(* IEC 61131-3 sources: PLC-IsaVODE/PLC-IsaVODE/samples/plc-programs (part 5) *)

(* ---- 533-TP_1.ST ---- *)
FUNCTION UDINT_TO_TIME2:TIME

	VAR_INPUT
		IN :	UDINT;
	END_VAR

	UDINT_TO_TIME2 := DINT_TO_TIME(UDINT_TO_DINT(IN));

END_FUNCTION

FUNCTION_BLOCK T_PLC_MS_block
	VAR_OUTPUT
		T_PLC_MS :	UDINT;
	END_VAR

	VAR_EXTERNAL
		PLC_TICKS_PER_SEC :	INT;
		PLC_SYS_TICK_CNT :	DINT;
	END_VAR

	VAR
		debug :	BOOL;(*Debug-Mode ON / OFF*)
		N :	INT;(*Debug-Faktor*)
		Offset :	UDINT;(*Debug-Offset*)
		temp :	DWORD := DWORD#1;(*Debug-Offset*)
		mode :	BOOL;(*modus*)
		faktor :	UDINT;(*Systemtakt-Faktor*)
		init :	BOOL;
		v_plc_ticks_per_sec :	UDINT;
		base :	UDINT := UDINT#1000;
	END_VAR

	IF init = FALSE THEN
		v_plc_ticks_per_sec := INT_TO_UDINT(PLC_TICKS_PER_SEC);
		IF v_plc_ticks_per_sec = UDINT#1024 THEN
			faktor := UDINT#1;
			mode := FALSE;
		ELSIF v_plc_ticks_per_sec > UDINT#0 THEN
			IF v_plc_ticks_per_sec <= base THEN
				faktor := base / v_plc_ticks_per_sec;
				mode := FALSE;
			ELSE
				faktor := v_plc_ticks_per_sec / base;
				mode := TRUE;
			END_IF;
		ELSE
			faktor := UDINT#1;
		END_IF;
		init := TRUE;
	END_IF;

	IF mode THEN
		T_PLC_MS := DINT_TO_UDINT(PLC_SYS_TICK_CNT) / faktor;
	ELSE
		T_PLC_MS := DINT_TO_UDINT(PLC_SYS_TICK_CNT) * faktor;
	END_IF;

	IF debug THEN
		T_PLC_MS := (DWORD_TO_UDINT(SHL(UDINT_TO_DWORD(T_PLC_MS),N) OR SHL(temp,N)) - UDINT#1) + Offset;
	END_IF;

END_FUNCTION_BLOCK

FUNCTION_BLOCK TP_1

	VAR_INPUT
		IN :	BOOL;
		PT :	TIME;
		RST :	BOOL;
	END_VAR

	VAR_OUTPUT
		Q :	BOOL;
	END_VAR

	VAR
		tx :	TIME;
		start :	TIME;
		ix :	BOOL;
		T_PLC_MS :	T_PLC_MS_block;
	END_VAR

	T_PLC_MS();
	tx := UDINT_TO_TIME(T_PLC_MS.T_PLC_MS);

	IF RST THEN
		Q := FALSE;
	ELSIF IN AND NOT ix THEN
		Q := TRUE;
		start := tx;
	ELSIF tx - start >= PT THEN
		Q := FALSE;
	END_IF;

	ix:= IN;

END_FUNCTION_BLOCK

PROGRAM program0
  VAR
	IN :	BOOL;
	PT :	TIME;
	RST :	BOOL;
	Q :	BOOL;
	func_block : TP_1;
  END_VAR
	func_block.IN  :=IN;
	func_block.PT  :=PT;
	func_block.RST  :=RST;
	func_block();
	Q := func_block.Q;
END_PROGRAM

CONFIGURATION Config0
	VAR_GLOBAL
		PLC_TICKS_PER_SEC :	INT;
		PLC_SYS_TICK_CNT :	DINT;
	END_VAR
	RESOURCE Res0 ON PLC
		TASK task0(INTERVAL := T#20ms,PRIORITY := 0);
		PROGRAM instance0 WITH task0 : program0;
	END_RESOURCE
END_CONFIGURATION

(* ---- 534-IRTRANS_RCV_8.ST ---- *)
FUNCTION_BLOCK IRTRANS_RCV_8_Block

	VAR_INPUT
		CMD :	BOOL;
	END_VAR

	VAR_IN_OUT
		DEV :	STRING;
		KEY :	STRING;
	END_VAR

	VAR_INPUT
		DEV_CODE :	STRING;
		KEY_CODE_0 :	STRING;
		KEY_CODE_1 :	STRING;
		KEY_CODE_2 :	STRING;
		KEY_CODE_3 :	STRING;
		KEY_CODE_4 :	STRING;
		KEY_CODE_5 :	STRING;
		KEY_CODE_6 :	STRING;
		KEY_CODE_7 :	STRING;
	END_VAR

	VAR_OUTPUT
		Q0 :	BOOL;
		Q1 :	BOOL;
		Q2 :	BOOL;
		Q3 :	BOOL;
		Q4 :	BOOL;
		Q5 :	BOOL;
		Q6 :	BOOL;
		Q7 :	BOOL;
	END_VAR

	VAR
		decode :	BOOL;
	END_VAR

	decode := cmd AND EQ_STRING(dev_code,dev);

	Q0 := EQ_STRING(key,key_code_0) AND decode;
	Q1 := EQ_STRING(key,key_code_1) AND decode;
	Q2 := EQ_STRING(key,key_code_2) AND decode;
	Q3 := EQ_STRING(key,key_code_3) AND decode;
	Q4 := EQ_STRING(key,key_code_4) AND decode;
	Q5 := EQ_STRING(key,key_code_5) AND decode;
	Q6 := EQ_STRING(key,key_code_6) AND decode;
	Q7 := EQ_STRING(key,key_code_7) AND decode;

END_FUNCTION_BLOCK

PROGRAM program0
	VAR
		CMD :	BOOL;
		DEV :	STRING;
		KEY :	STRING;
		DEV_CODE :	STRING;
		KEY_CODE_0 :	STRING;
		KEY_CODE_1 :	STRING;
		KEY_CODE_2 :	STRING;
		KEY_CODE_3 :	STRING;
		KEY_CODE_4 :	STRING;
		KEY_CODE_5 :	STRING;
		KEY_CODE_6 :	STRING;
		KEY_CODE_7 :	STRING;
		Q0 :	BOOL;
		Q1 :	BOOL;
		Q2 :	BOOL;
		Q3 :	BOOL;
		Q4 :	BOOL;
		Q5 :	BOOL;
		Q6 :	BOOL;
		Q7 :	BOOL;

		func_block : IRTRANS_RCV_8_Block;
	END_VAR
	func_block.CMD := CMD;
	func_block.DEV := DEV;
	func_block.KEY := KEY;
	func_block.DEV_CODE := DEV_CODE;
	func_block.KEY_CODE_0 := KEY_CODE_0;
	func_block.KEY_CODE_1 := KEY_CODE_1;
	func_block.KEY_CODE_2 := KEY_CODE_2;
	func_block.KEY_CODE_3 := KEY_CODE_3;
	func_block.KEY_CODE_4 := KEY_CODE_4;
	func_block.KEY_CODE_5 := KEY_CODE_5;
	func_block.KEY_CODE_6 := KEY_CODE_6;
	func_block.KEY_CODE_7 := KEY_CODE_7;

	func_block();
	DEV  := func_block.DEV;
	KEY  := func_block.KEY;
	Q0  := func_block.Q0;
	Q1  := func_block.Q1;
	Q2  := func_block.Q2;
	Q3  := func_block.Q3;
	Q4  := func_block.Q4;
	Q5  := func_block.Q5;
	Q6  := func_block.Q6;
	Q7  := func_block.Q7;

END_PROGRAM

CONFIGURATION Config0

  	RESOURCE Res0 ON PLC
    	TASK task0(INTERVAL := T#20ms,PRIORITY := 0);
    	PROGRAM instance0 WITH task0 : program0;
  	END_RESOURCE

END_CONFIGURATION

(* ---- 535-TP_X.ST ---- *)
FUNCTION UDINT_TO_TIME2:TIME

	VAR_INPUT
		IN :	UDINT;
	END_VAR

	UDINT_TO_TIME2 := DINT_TO_TIME(UDINT_TO_DINT(IN));

END_FUNCTION

FUNCTION_BLOCK T_PLC_MS_block
	VAR_OUTPUT
		T_PLC_MS :	UDINT;
	END_VAR

	VAR_EXTERNAL
		PLC_TICKS_PER_SEC :	INT;
		PLC_SYS_TICK_CNT :	DINT;
	END_VAR

	VAR
		debug :	BOOL;(*Debug-Mode ON / OFF*)
		N :	INT;(*Debug-Faktor*)
		Offset :	UDINT;(*Debug-Offset*)
		temp :	DWORD := DWORD#1;(*Debug-Offset*)
		mode :	BOOL;(*modus*)
		faktor :	UDINT;(*Systemtakt-Faktor*)
		init :	BOOL;
		v_plc_ticks_per_sec :	UDINT;
		base :	UDINT := UDINT#1000;
	END_VAR

	IF init = FALSE THEN
		v_plc_ticks_per_sec := INT_TO_UDINT(PLC_TICKS_PER_SEC);
		IF v_plc_ticks_per_sec = UDINT#1024 THEN
			faktor := UDINT#1;
			mode := FALSE;
		ELSIF v_plc_ticks_per_sec > UDINT#0 THEN
			IF v_plc_ticks_per_sec <= base THEN
				faktor := base / v_plc_ticks_per_sec;
				mode := FALSE;
			ELSE
				faktor := v_plc_ticks_per_sec / base;
				mode := TRUE;
			END_IF;
		ELSE
			faktor := UDINT#1;
		END_IF;
		init := TRUE;
	END_IF;

	IF mode THEN
		T_PLC_MS := DINT_TO_UDINT(PLC_SYS_TICK_CNT) / faktor;
	ELSE
		T_PLC_MS := DINT_TO_UDINT(PLC_SYS_TICK_CNT) * faktor;
	END_IF;

	IF debug THEN
		T_PLC_MS := (DWORD_TO_UDINT(SHL(UDINT_TO_DWORD(T_PLC_MS),N) OR SHL(temp,N)) - UDINT#1) + Offset;
	END_IF;

END_FUNCTION_BLOCK

FUNCTION_BLOCK TP_X
	VAR_INPUT
		IN :	BOOL;
		PT :	TIME;
	END_VAR

	VAR_OUTPUT
		Q :	BOOL;
		ET :	TIME;
	END_VAR

	VAR
		edge :	BOOL;
		start :	TIME;
		tx :	TIME;
		T_PLC_MS :	T_PLC_MS_block;
	END_VAR

	T_PLC_MS();
	tx := UDINT_TO_TIME2(T_PLC_MS.T_PLC_MS);

	IF IN AND NOT edge THEN
		start := tx;
		Q := PT > t#0ms;
	ELSIF Q THEN
		ET := tx - start;
		IF ET >= PT THEN
			Q := FALSE;
			ET := t#0ms;
		END_IF;
	END_IF;
	edge := IN;

END_FUNCTION_BLOCK

PROGRAM program0
  VAR
	IN :	BOOL;
	PT :	TIME;
	Q :	BOOL;
	ET :	TIME;
	func_block : TP_X;
  END_VAR
	func_block.IN  :=IN;
	func_block.PT  :=PT ;
	func_block();
	Q := func_block.Q;
	ET := func_block.ET;
END_PROGRAM

CONFIGURATION Config0
	VAR_GLOBAL
		PLC_TICKS_PER_SEC :	INT;
		PLC_SYS_TICK_CNT :	DINT;
	END_VAR
	RESOURCE Res0 ON PLC
		TASK task0(INTERVAL := T#20ms,PRIORITY := 0);
		PROGRAM instance0 WITH task0 : program0;
	END_RESOURCE
END_CONFIGURATION

(* ---- 536-EXEC.ST ---- *)
FUNCTION_BLOCK EXEC_Block
	VAR_INPUT
		STR :	STRING;
	END_VAR

	VAR_OUTPUT
		EXEC :	STRING;
	END_VAR

	VAR
		pos :	INT;
		R1 :	REAL;
		R2 :	REAL;
		operator :	STRING;
		temp :	STRING;
		uppercase :	uppercase;
		trim :	trim;
		findB_num :	findB_num;
		findB_nonum :	findB_nonum;
	END_VAR

	trim(str:=str);
	temp:=trim.trim;

	uppercase(str:=temp);
	exec:=uppercase.uppercase;

	findB_nonum(str:=exec);
	pos :=findB_nonum.findB_nonum;

	IF pos > 1 THEN
	temp := LEFT(EXEC,pos-1);
	findB_num(str:=temp);
	IF findB_num.findB_num > 0 THEN
	R1 := STRING_TO_REAL(temp);
	END_IF;
	END_IF;
	temp := RIGHT(exec,LEN(exec)-pos);
	R2 := STRING_TO_REAL(temp);
	exec := LEFT(exec,pos);

	findB_num(str:=exec);
	pos :=findB_num.findB_num;
	operator := RIGHT(exec,LEN(exec) - pos);
	IF EQ_STRING(operator,'') AND LEN(str) = 0 THEN
		exec := '';
		RETURN;
	ELSIF EQ_STRING(operator,'') THEN
		exec := str;
		RETURN;
	END_IF;
	IF EQ_STRING(operator,'^') THEN
		exec := REAL_TO_STRING(EXPT(R1, R2),'%f');
	ELSIF EQ_STRING(operator,'SQRT') THEN
		exec := REAL_TO_STRING(SQRT(R2),'%f');
	ELSIF EQ_STRING(operator,'SIN') THEN
		exec := REAL_TO_STRING(SIN(r2),'%f');
	ELSIF EQ_STRING(operator,'COS') THEN
		exec := REAL_TO_STRING(COS(r2),'%f');
	ELSIF EQ_STRING(operator,'TAN') THEN
		exec := REAL_TO_STRING(TAN(R2),'%f');
	ELSIF EQ_STRING(operator,'*') THEN
		exec := REAL_TO_STRING(R1 * R2,'%f');
	ELSIF EQ_STRING(operator,'/') THEN
		IF R2 <> 0.0 THEN exec := REAL_TO_STRING(R1 / R2,'%f'); ELSE exec := 'ERROR'; END_IF;
	ELSIF EQ_STRING(operator,'+') THEN
		exec := REAL_TO_STRING(r1 + r2,'%f');
	ELSIF EQ_STRING(operator,'-') THEN
		exec := REAL_TO_STRING(r1 - r2,'%f');
	ELSE
		exec := 'ERROR';
	END_IF;
	IF EQ_STRING(EXEC,'ERROR') THEN
		RETURN;
	ELSIF FIND(EXEC,'.') = 0 THEN
		EXEC := CONCAT(EXEC, '.0');
	ELSE
	temp := RIGHT(EXEC,1);
	IF EQ_STRING(temp,'.') THEN
		EXEC := CONCAT(EXEC,'0');
	END_IF;
	END_IF;

END_FUNCTION_BLOCK

PROGRAM program0
	VAR
		STR :	STRING;

		EXEC :	STRING;

		func_block : EXEC_Block;
	END_VAR
	func_block.STR := STR;
	func_block();
	EXEC  := func_block.EXEC;
END_PROGRAM

CONFIGURATION Config0
	RESOURCE Res0 ON PLC
		TASK task0(INTERVAL := T#20ms,PRIORITY := 0);
		PROGRAM instance0 WITH task0 : program0;
	END_RESOURCE
END_CONFIGURATION

(* ---- 537-FILE_BLOCK.ST ---- *)
TYPE
  oscat_FILE_SERVER_DATA : STRUCT
	FILE_OPEN	: BOOL;
    FILENAME 	: STRING;
    MODE	 	: BYTE;
    OFFSET   	: UDINT;
    FILE_SIZE   : UDINT;
    AUTO_CLOSE	: TIME;
    ERROR	 	: BYTE;
  END_STRUCT;

  oscat_NW_BUF_LONG  : ARRAY [0..4095] OF BYTE;
  oscat_NETWORK_BUFFER :
  STRUCT
    SIZE   : UINT;
    BUFFER : oscat_NW_BUF_LONG;
  END_STRUCT;
END_TYPE

FUNCTION_BLOCK FILE_BLOCK

	VAR_IN_OUT
		MODE :	BYTE;
		FILENAME :	STRING;
		FSD :	oscat_FILE_SERVER_DATA;
		PT :	oscat_NETWORK_BUFFER;
	END_VAR

	VAR_INPUT
		POS :	UDINT;
	END_VAR

	VAR_OUTPUT
		ERROR :	BYTE;
		DATA :	BYTE;
	END_VAR

	VAR
		stepp :	INT;
		i :	INT;
		data_start :	UDINT;
		data_stop :	UDINT;
	END_VAR

	CASE stepp OF
	0:	IF MODE > BYTE#0 THEN
			ERROR := BYTE#0;
			IF FSD.FILE_OPEN AND (FSD.FILE_SIZE = UDINT#0 OR POS >= FSD.FILE_SIZE) THEN
				ERROR := BYTE#255;
				MODE := BYTE#0;
			ELSIF POS < data_start OR POS > data_stop OR NOT FSD.FILE_OPEN THEN
				FSD.FILENAME := FILENAME;
				FSD.MODE := BYTE#1;
				FSD.OFFSET := POS;
				PT.SIZE := UINT#65535;
				data_start := UDINT#0;
				data_stop := UDINT#0;
				stepp := 10;
			ELSE
				i := UDINT_TO_INT(POS - data_start);
				DATA := PT.BUFFER[i];
				MODE := BYTE#0;
			END_IF;
		END_IF;

	10:	IF FSD.MODE = BYTE#0 THEN
			IF FSD.ERROR > BYTE#0 THEN
				ERROR := FSD.ERROR;
				MODE := BYTE#0;
			ELSE
				data_start := POS;
				data_stop := POS + UINT_TO_UDINT(PT.SIZE) - UDINT#1;
			END_IF;
			stepp := 0;
		END_IF;
	END_CASE;
END_FUNCTION_BLOCK

PROGRAM program0
	VAR
		MODE :	BYTE;
		FILENAME :	STRING;
		FSD :	oscat_FILE_SERVER_DATA;
		PT :	oscat_NETWORK_BUFFER;
		POS :	UDINT;
		ERROR :	BYTE;
		DATA :	BYTE;

		func_block : FILE_BLOCK;
	END_VAR
	func_block.MODE    :=MODE    ;
	func_block.FILENAME:=FILENAME;
	func_block.FSD     :=FSD     ;
	func_block.PT      :=PT      ;
	func_block.POS     :=POS     ;
	func_block();
	MODE    := func_block.MODE    ;
	FILENAME:= func_block.FILENAME;
	FSD     := func_block.FSD     ;
	PT      := func_block.PT      ;
	ERROR   := func_block.ERROR;
	DATA    := func_block.DATA;

END_PROGRAM

CONFIGURATION Config0
  RESOURCE Res0 ON PLC
    TASK task0(INTERVAL := T#20ms,PRIORITY := 0);
    PROGRAM instance0 WITH task0 : program0;
  END_RESOURCE
END_CONFIGURATION

(* ---- 538-TMAX.ST ---- *)
FUNCTION UDINT_TO_TIME2:TIME

	VAR_INPUT
		IN :	UDINT;
	END_VAR

	UDINT_TO_TIME2 := DINT_TO_TIME(UDINT_TO_DINT(IN));

END_FUNCTION

FUNCTION_BLOCK T_PLC_MS_block
	VAR_OUTPUT
		T_PLC_MS :	UDINT;
	END_VAR

	VAR_EXTERNAL
		PLC_TICKS_PER_SEC :	INT;
		PLC_SYS_TICK_CNT :	DINT;
	END_VAR

	VAR
		debug :	BOOL;(*Debug-Mode ON / OFF*)
		N :	INT;(*Debug-Faktor*)
		Offset :	UDINT;(*Debug-Offset*)
		temp :	DWORD := DWORD#1;(*Debug-Offset*)
		mode :	BOOL;(*modus*)
		faktor :	UDINT;(*Systemtakt-Faktor*)
		init :	BOOL;
		v_plc_ticks_per_sec :	UDINT;
		base :	UDINT := UDINT#1000;
	END_VAR

	IF init = FALSE THEN
		v_plc_ticks_per_sec := INT_TO_UDINT(PLC_TICKS_PER_SEC);
		IF v_plc_ticks_per_sec = UDINT#1024 THEN
			faktor := UDINT#1;
			mode := FALSE;
		ELSIF v_plc_ticks_per_sec > UDINT#0 THEN
			IF v_plc_ticks_per_sec <= base THEN
				faktor := base / v_plc_ticks_per_sec;
				mode := FALSE;
			ELSE
				faktor := v_plc_ticks_per_sec / base;
				mode := TRUE;
			END_IF;
		ELSE
			faktor := UDINT#1;
		END_IF;
		init := TRUE;
	END_IF;

	IF mode THEN
		T_PLC_MS := DINT_TO_UDINT(PLC_SYS_TICK_CNT) / faktor;
	ELSE
		T_PLC_MS := DINT_TO_UDINT(PLC_SYS_TICK_CNT) * faktor;
	END_IF;

	IF debug THEN
		T_PLC_MS := (DWORD_TO_UDINT(SHL(UDINT_TO_DWORD(T_PLC_MS),N) OR SHL(temp,N)) - UDINT#1) + Offset;
	END_IF;

END_FUNCTION_BLOCK

FUNCTION_BLOCK TMAX

	VAR_INPUT
		IN :	BOOL;
		PT :	TIME;
	END_VAR

	VAR_OUTPUT
		Q :	BOOL;
		Z :	BOOL;
	END_VAR

	VAR
		tx :	TIME;
		start :	TIME;
		last_in :	BOOL;
		T_PLC_MS :	T_PLC_MS_block;
	END_VAR

	T_PLC_MS();
	tx:= UDINT_TO_TIME(T_PLC_MS.T_PLC_MS);

	Z := FALSE;

	IF NOT in THEN
		Q := FALSE;
	ELSIF IN AND NOT last_in THEN
		Q := TRUE;
		start := tx;
	ELSIF (tx - start >= PT) AND Q THEN
		Q := FALSE;
		Z := TRUE;
	END_IF;

	last_in := IN;

END_FUNCTION_BLOCK

PROGRAM program0
  VAR
	IN :	BOOL;
	PT :	TIME;
	Q :	BOOL;
	Z :	BOOL;
	func_block : TMAX;
  END_VAR
	func_block.IN  :=IN;
	func_block.PT  :=PT;
	func_block();
	Q := func_block.Q;
	Z := func_block.Z;

END_PROGRAM

CONFIGURATION Config0
	VAR_GLOBAL
		PLC_TICKS_PER_SEC :	INT;
		PLC_SYS_TICK_CNT :	DINT;
	END_VAR
	RESOURCE Res0 ON PLC
		TASK task0(INTERVAL := T#20ms,PRIORITY := 0);
		PROGRAM instance0 WITH task0 : program0;
	END_RESOURCE
END_CONFIGURATION

(* ---- 539-M_T.ST ---- *)
FUNCTION_BLOCK T_PLC_MS_block
	VAR_OUTPUT
		T_PLC_MS :	UDINT;
	END_VAR

	VAR_EXTERNAL
		PLC_TICKS_PER_SEC :	INT;
		PLC_SYS_TICK_CNT :	DINT;
	END_VAR

	VAR
		debug :	BOOL;(*Debug-Mode ON / OFF*)
		N :	INT;(*Debug-Faktor*)
		Offset :	UDINT;(*Debug-Offset*)
		temp :	DWORD := DWORD#1;(*Debug-Offset*)
		mode :	BOOL;(*modus*)
		faktor :	UDINT;(*Systemtakt-Faktor*)
		init :	BOOL;
		v_plc_ticks_per_sec :	UDINT;
		base :	UDINT := UDINT#1000;
	END_VAR

	IF init = FALSE THEN
		v_plc_ticks_per_sec := INT_TO_UDINT(PLC_TICKS_PER_SEC);
		IF v_plc_ticks_per_sec = UDINT#1024 THEN
			faktor := UDINT#1;
			mode := FALSE;
		ELSIF v_plc_ticks_per_sec > UDINT#0 THEN
			IF v_plc_ticks_per_sec <= base THEN
				faktor := base / v_plc_ticks_per_sec;
				mode := FALSE;
			ELSE
				faktor := v_plc_ticks_per_sec / base;
				mode := TRUE;
			END_IF;
		ELSE
			faktor := UDINT#1;
		END_IF;
		init := TRUE;
	END_IF;

	IF mode THEN
		T_PLC_MS := DINT_TO_UDINT(PLC_SYS_TICK_CNT) / faktor;
	ELSE
		T_PLC_MS := DINT_TO_UDINT(PLC_SYS_TICK_CNT) * faktor;
	END_IF;

	IF debug THEN
		T_PLC_MS := (DWORD_TO_UDINT(SHL(UDINT_TO_DWORD(T_PLC_MS),N) OR SHL(temp,N)) - UDINT#1) + Offset;
	END_IF;
END_FUNCTION_BLOCK

FUNCTION_BLOCK M_T_Block

	VAR_INPUT
		IN :	BOOL;
		TMAX :	TIME := t#10d;
		RST :	BOOL;
	END_VAR

	VAR_OUTPUT
		PT :	TIME;
		ET :	TIME;
	END_VAR

	VAR
		edge :	BOOL;
		start :	TIME;
		tx :	TIME;
		T_PLC_MS :	T_PLC_MS_Block;
	END_VAR

	(*@KEY@: WORKSHEET
	NAME: M_T
	IEC_LANGUAGE: ST
	*)
	(* read system timer *)
	T_PLC_MS();
	tx:= UDINT_TO_TIME(T_PLC_MS.T_PLC_MS);

	IF RST OR ET >= TMAX THEN
		PT := t#0s;
		ET := PT;
	ELSIF IN THEN
		IF NOT edge THEN start := tx; END_IF;
		ET := tx - start;
	ELSE
		PT := ET;
	END_IF;
	edge := IN;

END_FUNCTION_BLOCK

PROGRAM program0

	VAR
		IN :	BOOL;
		TMAX :	TIME := t#10d;
		RST :	BOOL;

		PT :	TIME;
		ET :	TIME;

		func_block : M_T_Block;
	END_VAR
	func_block.IN := IN;
	func_block.TMAX := TMAX;
	func_block.RST := RST;

	func_block();
	PT := func_block.PT;
	ET := func_block.ET;

END_PROGRAM

CONFIGURATION Config0

	VAR_GLOBAL
		PLC_TICKS_PER_SEC :	INT;
		PLC_SYS_TICK_CNT :	DINT;
	END_VAR

	RESOURCE Res0 ON PLC
		TASK task0(INTERVAL := T#20ms,PRIORITY := 0);
		PROGRAM instance0 WITH task0 : program0;
	END_RESOURCE

END_CONFIGURATION

(* ---- 540-FT_IMP.ST ---- *)
FUNCTION_BLOCK T_PLC_US_Block

	VAR_OUTPUT
		T_PLC_US :	UDINT;
	END_VAR

	VAR_EXTERNAL
		PLC_TICKS_PER_SEC :	INT;
		PLC_SYS_TICK_CNT :	DINT;
	END_VAR

	VAR
		debug :	BOOL;
		N :	INT;
		Offset :	UDINT;
		temp :	DWORD := DWORD#1;
		mode :	BOOL;
		faktor :	UDINT;
		init :	BOOL;
		v_plc_ticks_per_sec :	UDINT;
		base :	UDINT := UDINT#1000000;
	END_VAR

	IF init = FALSE THEN
		v_plc_ticks_per_sec := INT_TO_UDINT(PLC_TICKS_PER_SEC);
		IF v_plc_ticks_per_sec = UDINT#1024 THEN
			faktor := UDINT#1000;
			mode := FALSE;
		ELSIF v_plc_ticks_per_sec > UDINT#0 THEN
			IF v_plc_ticks_per_sec <= base THEN
				faktor := base / v_plc_ticks_per_sec;
				mode := FALSE;
			ELSE
				faktor := v_plc_ticks_per_sec / base;
				mode := TRUE;
			END_IF;
		ELSE
			faktor := UDINT#1;
		END_IF;
		init := TRUE;
	END_IF;

	IF mode THEN
		T_PLC_US := DINT_TO_UDINT(PLC_SYS_TICK_CNT) / faktor;
	ELSE
		T_PLC_US := DINT_TO_UDINT(PLC_SYS_TICK_CNT) * faktor;
	END_IF;

	IF debug THEN
		T_PLC_US := (DWORD_TO_UDINT(SHL(UDINT_TO_DWORD(T_PLC_US),N) OR SHL(temp,N)) - UDINT#1) + Offset;
	END_IF;

END_FUNCTION_BLOCK

FUNCTION_BLOCK FT_PT1

	VAR_INPUT
		IN :	REAL;
		T :	TIME;
		K :	REAL := 1.0;
	END_VAR

	VAR_OUTPUT
		OUT :	REAL;
	END_VAR

	VAR
		last :	UDINT;
		tx :	UDINT;
		init :	BOOL;
		T_PLC_US :	T_PLC_US_Block;
	END_VAR

	T_PLC_US();
	tx:= T_PLC_US.T_PLC_US;

	IF NOT init OR T = t#0s THEN
		init := TRUE;
		out := K * in;
	ELSE
		out := out + (in * K - out) * UDINT_TO_REAL(Tx - last) / TIME_TO_REAL(T) * 1.0E-3;
		IF ABS(out) < 1.0E-20 THEN out := 0.0; END_IF;
	END_IF;
	last := tx;

END_FUNCTION_BLOCK

FUNCTION_BLOCK FT_IMP

	VAR_INPUT
		IN :	REAL;
		T :	TIME;
		K :	REAL := 1.0;
	END_VAR

	VAR_OUTPUT
		OUT :	REAL;
	END_VAR

	VAR
		t1 :	FT_PT1;
	END_VAR

	T1(in:= in, T:=T);
	out := (in - t1.out) * K;

END_FUNCTION_BLOCK

PROGRAM program0
  VAR
	IN :	REAL;
	T :	TIME;
	K :	REAL;

	OUT :	REAL;

	func_block : FT_IMP;
  END_VAR
	func_block.IN :=IN ;
	func_block.T  :=T  ;
	func_block.K  :=K  ;
	func_block();
	OUT := func_block.OUT;
END_PROGRAM

CONFIGURATION Config0

	VAR_GLOBAL
		PLC_TICKS_PER_SEC :	INT;
		PLC_SYS_TICK_CNT :	DINT;
	END_VAR

	RESOURCE Res0 ON PLC
		TASK task0(INTERVAL := T#20ms,PRIORITY := 0);
		PROGRAM instance0 WITH task0 : program0;
	END_RESOURCE

END_CONFIGURATION

(* ---- 541-NET_VAR_BUFFER.ST ---- *)
TYPE
	oscat_aB1_64 : ARRAY[1..64] OF BYTE;
END_TYPE

TYPE

	oscat_NW_BUF_LONG  : ARRAY [0..4095] OF BYTE;

	oscat_NETWORK_BUFFER :
	STRUCT
		SIZE   : UINT;
		BUFFER : oscat_NW_BUF_LONG;
	END_STRUCT;

END_TYPE

TYPE oscat_NET_VAR_DATA :
	STRUCT
		CYCLE : UDINT;
		STATE : BYTE;
		INDEX : INT;
		ID_MAX : USINT;
		ERROR_ID : BYTE;
		BUF_SIZE : UINT;
		S_BUF : oscat_NETWORK_BUFFER;
		R_BUF : oscat_NETWORK_BUFFER;
	END_STRUCT;
END_TYPE

FUNCTION_BLOCK NET_VAR_BUFFER_Block

	VAR_OUTPUT
		ID :	BYTE;
	END_VAR

	VAR_IN_OUT
		BUF_IN :	oscat_aB1_64;
		BUF_OUT :	oscat_aB1_64;
		X :	oscat_NET_VAR_DATA;
	END_VAR

	VAR
		size :	INT;
		init :	BOOL;
		index :	INT;
		index2 :	INT;
	END_VAR

	IF NOT init THEN
		init := TRUE;
		X.ID_MAX := X.ID_MAX + USINT#1;
		ID := USINT_TO_BYTE(X.ID_MAX);
	END_IF;

	IF X.STATE > BYTE#0 AND X.ERROR_ID = BYTE#0 THEN
		index := X.index;
		IF X.STATE = BYTE#1 THEN
			size := 64;
			IF INT_TO_UINT(index + 3 + size) > X.BUF_SIZE THEN
				X.ERROR_ID := ID;
			ELSE
				X.S_BUF.BUFFER[index] := ID;
				index := index + 1;
				X.S_BUF.BUFFER[index] := BYTE#20;
				index := index + 1;
				X.S_BUF.BUFFER[index] := INT_TO_BYTE(size);
				index := index + 1;
				FOR index2 := 1 TO size DO
					X.S_BUF.BUFFER[index] := BUF_IN[index2];
					index := index + 1;
				END_FOR;
			END_IF;
		ELSIF X.STATE = BYTE#2 THEN
			index2 := index + 1;
			IF X.R_BUF.BUFFER[index] <> ID OR X.R_BUF.BUFFER[index2] <> BYTE#20 THEN
				X.ERROR_ID := ID;
			ELSE
				index := index + 2;
				size := BYTE_TO_INT(X.R_BUF.BUFFER[index]);
				index := index + 1;
				FOR index2 := 1 TO size DO
					BUF_OUT[index2] := X.R_BUF.BUFFER[index];
					index := index + 1;
				END_FOR;
			END_IF;
		END_IF;
		X.index := index;
	END_IF;

END_FUNCTION_BLOCK

PROGRAM program0
	VAR
		BUF_IN :	oscat_aB1_64;
		BUF_OUT :	oscat_aB1_64;
		X :	oscat_NET_VAR_DATA;
		ID :	BYTE;

		func_block : NET_VAR_BUFFER_Block;
	END_VAR
	func_block.BUF_IN := BUF_IN;
	func_block.BUF_OUT := BUF_OUT;
	func_block.X := X;

	func_block();
  	BUF_IN  := func_block.BUF_IN;
	BUF_OUT  := func_block.BUF_OUT;
	X  := func_block.X;
	ID  := func_block.ID;

END_PROGRAM

CONFIGURATION Config0
	RESOURCE Res0 ON PLC
		TASK task0(INTERVAL := T#20ms,PRIORITY := 0);
		PROGRAM instance0 WITH task0 : program0;
	END_RESOURCE
END_CONFIGURATION

(* ---- 542-GEN_PULSE.ST ---- *)
FUNCTION UDINT_TO_TIME2:TIME

	VAR_INPUT
		IN :	UDINT;
	END_VAR

	UDINT_TO_TIME2 := DINT_TO_TIME(UDINT_TO_DINT(IN));

END_FUNCTION

FUNCTION_BLOCK T_PLC_MS_block
	VAR_OUTPUT
		T_PLC_MS :	UDINT;
	END_VAR

	VAR_EXTERNAL
		PLC_TICKS_PER_SEC :	INT;
		PLC_SYS_TICK_CNT :	DINT;
	END_VAR

	VAR
		debug :	BOOL;(*Debug-Mode ON / OFF*)
		N :	INT;(*Debug-Faktor*)
		Offset :	UDINT;(*Debug-Offset*)
		temp :	DWORD := DWORD#1;(*Debug-Offset*)
		mode :	BOOL;(*modus*)
		faktor :	UDINT;(*Systemtakt-Faktor*)
		init :	BOOL;
		v_plc_ticks_per_sec :	UDINT;
		base :	UDINT := UDINT#1000;
	END_VAR

	IF init = FALSE THEN
		v_plc_ticks_per_sec := INT_TO_UDINT(PLC_TICKS_PER_SEC);
		IF v_plc_ticks_per_sec = UDINT#1024 THEN
			faktor := UDINT#1;
			mode := FALSE;
		ELSIF v_plc_ticks_per_sec > UDINT#0 THEN
			IF v_plc_ticks_per_sec <= base THEN
				faktor := base / v_plc_ticks_per_sec;
				mode := FALSE;
			ELSE
				faktor := v_plc_ticks_per_sec / base;
				mode := TRUE;
			END_IF;
		ELSE
			faktor := UDINT#1;
		END_IF;
		init := TRUE;
	END_IF;

	IF mode THEN
		T_PLC_MS := DINT_TO_UDINT(PLC_SYS_TICK_CNT) / faktor;
	ELSE
		T_PLC_MS := DINT_TO_UDINT(PLC_SYS_TICK_CNT) * faktor;
	END_IF;

	IF debug THEN
		T_PLC_MS := (DWORD_TO_UDINT(SHL(UDINT_TO_DWORD(T_PLC_MS),N) OR SHL(temp,N)) - UDINT#1) + Offset;
	END_IF;

END_FUNCTION_BLOCK

FUNCTION_BLOCK GEN_PULSE_Block

	VAR_INPUT
		ENQ :	BOOL := TRUE;
		PTH :	TIME;
		PTL :	TIME;
	END_VAR

	VAR_OUTPUT
		Q :	BOOL;
	END_VAR

	VAR
		T_PLC_MS :	T_PLC_MS_block;
		tx :	TIME;
		tn :	TIME;
		init :	BOOL;
	END_VAR

	IF enq THEN
		T_PLC_MS();
		tx:= UDINT_TO_TIME(T_PLC_MS.T_PLC_MS);
		IF NOT init THEN init := TRUE; tn := tx; END_IF;
		IF tx - tn >= SEL(Q, PTL, PTH) THEN
			tn := tn + SEL(Q, PTL, PTH);
			Q := NOT Q;
		END_IF;
	ELSE
		Q := FALSE;
		init := FALSE;
	END_IF;

END_FUNCTION_BLOCK

PROGRAM program0
  VAR
	ENQ :	BOOL := TRUE;
	PTH :	TIME;
	PTL :	TIME;
	Q :	BOOL;
	func_block : GEN_PULSE_Block;
  END_VAR
	func_block.ENQ  :=ENQ;
	func_block.PTH  :=PTH;
	func_block.PTL  :=PTL;
	func_block();
	Q := func_block.Q;

END_PROGRAM

CONFIGURATION Config0
	VAR_GLOBAL
		PLC_TICKS_PER_SEC :	INT;
		PLC_SYS_TICK_CNT :	DINT;
	END_VAR
	RESOURCE Res0 ON PLC
		TASK task0(INTERVAL := T#20ms,PRIORITY := 0);
		PROGRAM instance0 WITH task0 : program0;
	END_RESOURCE
END_CONFIGURATION

(* ---- 543-FT_DERIV.ST ---- *)
FUNCTION_BLOCK T_PLC_US_Block
	VAR_OUTPUT
		T_PLC_US :	UDINT;
	END_VAR

	VAR_EXTERNAL
		PLC_TICKS_PER_SEC :	INT;
		PLC_SYS_TICK_CNT :	DINT;
	END_VAR

	VAR
		debug :	BOOL;
		N :	INT;
		Offset :	UDINT;
		temp :	DWORD := DWORD#1;
		mode :	BOOL;
		faktor :	UDINT;
		init :	BOOL;
		v_plc_ticks_per_sec :	UDINT;
		base :	UDINT := UDINT#1000000;
	END_VAR

	IF init = FALSE THEN
		v_plc_ticks_per_sec := INT_TO_UDINT(PLC_TICKS_PER_SEC);
		IF v_plc_ticks_per_sec = UDINT#1024 THEN
			faktor := UDINT#1000;
			mode := FALSE;
		ELSIF v_plc_ticks_per_sec > UDINT#0 THEN
			IF v_plc_ticks_per_sec <= base THEN
				faktor := base / v_plc_ticks_per_sec;
				mode := FALSE;
			ELSE
				faktor := v_plc_ticks_per_sec / base;
				mode := TRUE;
			END_IF;
		ELSE
			faktor := UDINT#1;
		END_IF;
		init := TRUE;
	END_IF;

	IF mode THEN
		T_PLC_US := DINT_TO_UDINT(PLC_SYS_TICK_CNT) / faktor;
	ELSE
		T_PLC_US := DINT_TO_UDINT(PLC_SYS_TICK_CNT) * faktor;
	END_IF;

	IF debug THEN
		T_PLC_US := (DWORD_TO_UDINT(SHL(UDINT_TO_DWORD(T_PLC_US),N) OR SHL(temp,N)) - UDINT#1) + Offset;
	END_IF;
END_FUNCTION_BLOCK

FUNCTION_BLOCK FT_DERIV
	VAR_INPUT
		IN :	REAL;
		K :	REAL := 1.0;
		RUN :	BOOL := TRUE;
	END_VAR

	VAR_OUTPUT
		OUT :	REAL;
	END_VAR

	VAR
		old :	REAL;
		tx :	UDINT;
		last :	UDINT;
		init :	BOOL;
		tc :	REAL;
		T_PLC_US :	T_PLC_US_Block;
	END_VAR

	T_PLC_US();
	tx:= T_PLC_US.T_PLC_US;
	tc := UDINT_TO_REAL(tx - last);

	IF NOT init THEN
		init := TRUE;
		old := in;
	ELSIF run AND tc > 0.0 THEN
		out := (in - old) / tc * 1000000.0 * K;
		old := in;
	ELSE
		out := 0.0;
	END_IF;

	last := tx;

	T_PLC_US();
	tx:= T_PLC_US.T_PLC_US;

	IF NOT init THEN
		init := TRUE;
	ELSIF run AND tx - last > UDINT#0 THEN
		out := (in - old) / UDINT_TO_REAL(tx - last) * 1000000.0 * K;
	ELSE
		out := 0.0;
	END_IF;
	old := in;
	last := tx;
END_FUNCTION_BLOCK

PROGRAM program0
  VAR
	IN  :	REAL;
	K   :	REAL;
	RUN :	BOOL;

	OUT :	REAL;

	func_block : FT_DERIV;
  END_VAR
	func_block.IN :=IN ;
	func_block.K  :=K  ;
	func_block.RUN:=RUN;
	func_block();
	OUT := func_block.OUT;
END_PROGRAM

CONFIGURATION Config0
	VAR_GLOBAL
		PLC_TICKS_PER_SEC :	INT;
		PLC_SYS_TICK_CNT :	DINT;
	END_VAR

	RESOURCE Res0 ON PLC
		TASK task0(INTERVAL := T#20ms,PRIORITY := 0);
		PROGRAM instance0 WITH task0 : program0;
	END_RESOURCE
END_CONFIGURATION

(* ---- 544-REAL_TO_FRAC.ST ---- *)
TYPE oscat_FRACTION :
	STRUCT
		NUMERATOR : INT;
		DENOMINATOR : INT;
	END_STRUCT;
END_TYPE

FUNCTION_BLOCK REAL_TO_FRAC_Block

	VAR_INPUT
		X :	REAL;
		N :	INT;
	END_VAR

	VAR_OUTPUT
		REAL_TO_FRAC :	oscat_FRACTION;
	END_VAR

	VAR
		temp :	DINT;
		sign :	BOOL;
		X_gerundet :	DINT;
		X_ohne_Nachkomma :	REAL;
		Numerator :	DINT := 1;
		Denominator :	DINT := 0;
		Numerator_old :	DINT := 0;
		Denominator_old :	DINT := 1;
	END_VAR

	IF X < 0.0 THEN
		sign := TRUE;								(* Vorzeichen merken *)
		X := ABS(X);								(* Absolutwert berechnen *)
	END_IF;

	REPEAT
		X_gerundet := REAL_TO_DINT(X);

		temp := numerator * X_gerundet + numerator_old;		(* Zaehler um Vorkammawert erweitern *)
		numerator_old := numerator;							(* Zaehler der letzten Berechnung speichern *)
		numerator := temp;									(* Zaehler dieser Berechnung speichern *)

		temp := denominator * X_gerundet + denominator_old;	(* Nenner um Vorkammawert erweitern *)
		denominator_old := denominator;						(* Nenner der letzten Berechnung speichern *)
		denominator := temp;								(* Nenner dieser Berechnung speichern *)

		X_ohne_Nachkomma := DINT_TO_REAL(X_gerundet);
		IF X = X_ohne_Nachkomma THEN						(* Bruch geht ohne Rest auf *)
			IF ABS(denominator) <= INT_TO_DINT(N) THEN		(* kein Rundungsfehler *)
				numerator_old := numerator;					(* Numerator_old wird von Funktion zur�ckgegeben *)
				denominator_old := denominator;				(* Denominator_old wird von Funktion zur�ckgegeben *)
			END_IF;
			EXIT;											(* keine weitere Berechnung notwendig *)
		ELSE
			X := 1.0 / (X - X_ohne_Nachkomma);				(* Kehrwert vom Rest -> Neuer Bruch *)
		END_IF;

	UNTIL
		( ABS(Denominator) > INT_TO_DINT(N))
	END_REPEAT;

	IF sign THEN
		REAL_TO_FRAC.NUMERATOR := -1 * ABS(DINT_TO_INT(numerator_old));
	ELSE
		REAL_TO_FRAC.NUMERATOR :=  ABS(DINT_TO_INT(numerator_old));
	END_IF;

	REAL_TO_FRAC.DENOMINATOR := ABS(DINT_TO_INT(denominator_old));

END_FUNCTION_BLOCK

PROGRAM program0

	VAR
		X :	REAL;
		N :	INT;

        REAL_TO_FRAC :	oscat_FRACTION;
		func_block : REAL_TO_FRAC_Block;
	END_VAR
		func_block.X := X;
		func_block.N := N;
		func_block();
		REAL_TO_FRAC := func_block.REAL_TO_FRAC;

END_PROGRAM

CONFIGURATION Config0

	RESOURCE Res0 ON PLC
		TASK task0(INTERVAL := T#20ms,PRIORITY := 0);
		PROGRAM instance0 WITH task0 : program0;
	END_RESOURCE

END_CONFIGURATION

(* ---- 545-FT_TN8.ST ---- *)
TYPE
  	oscat_arr_0_7               : ARRAY [0..7]    OF REAL;
END_TYPE

FUNCTION_BLOCK T_PLC_MS_Block
	VAR_OUTPUT
		T_PLC_MS :	UDINT;
	END_VAR

	VAR_EXTERNAL
		PLC_TICKS_PER_SEC :	INT;
		PLC_SYS_TICK_CNT :	DINT;
	END_VAR

	VAR
		debug :	BOOL;(*Debug-Mode ON / OFF*)
		N :	INT;(*Debug-Faktor*)
		Offset :	UDINT;(*Debug-Offset*)
		temp :	DWORD := DWORD#1;(*Debug-Offset*)
		mode :	BOOL;(*modus*)
		faktor :	UDINT;(*Systemtakt-Faktor*)
		init :	BOOL;
		v_plc_ticks_per_sec :	UDINT;
		base :	UDINT := UDINT#1000;
	END_VAR

	IF init = FALSE THEN
		v_plc_ticks_per_sec := INT_TO_UDINT(PLC_TICKS_PER_SEC);
		IF v_plc_ticks_per_sec = UDINT#1024 THEN
			faktor := UDINT#1;
			mode := FALSE;
		ELSIF v_plc_ticks_per_sec > UDINT#0 THEN
			IF v_plc_ticks_per_sec <= base THEN
				faktor := base / v_plc_ticks_per_sec;
				mode := FALSE;
			ELSE
				faktor := v_plc_ticks_per_sec / base;
				mode := TRUE;
			END_IF;
		ELSE
			faktor := UDINT#1;
		END_IF;
		init := TRUE;
	END_IF;

	IF mode THEN
		T_PLC_MS := DINT_TO_UDINT(PLC_SYS_TICK_CNT) / faktor;
	ELSE
		T_PLC_MS := DINT_TO_UDINT(PLC_SYS_TICK_CNT) * faktor;
	END_IF;

	IF debug THEN
		T_PLC_MS := (DWORD_TO_UDINT(SHL(UDINT_TO_DWORD(T_PLC_MS),N) OR SHL(temp,N)) - UDINT#1) + Offset;
	END_IF;
END_FUNCTION_BLOCK

FUNCTION_BLOCK FT_TN8

	VAR_INPUT
		IN :	REAL;
		T :	TIME;
	END_VAR

	VAR_OUTPUT
		OUT :	REAL;
		TRIG :	BOOL;
	END_VAR

	VAR
		length :	INT := 8;
		X :	oscat_arr_0_7;
		cnt :	INT;
		last :	TIME;
		tx :	TIME;
		init :	BOOL;
		T_PLC_MS :	T_PLC_MS_Block;
	END_VAR

	T_PLC_MS();
	tx:= UDINT_TO_TIME(T_PLC_MS.T_PLC_MS);

	trig := FALSE;
	IF NOT init THEN
		x[cnt] := in;
		init := TRUE;
		last := tx;
	ELSIF tx - last >= (T / length) THEN
		IF cnt = length - 1 THEN cnt := 0; ELSE cnt := cnt + 1; END_IF;
		Out := X[cnt];
		x[cnt] := in;
		last := tx;
		trig := TRUE;
	END_IF;

END_FUNCTION_BLOCK

PROGRAM program0
  VAR
	IN :	REAL;
	T :	TIME;

	OUT :	REAL;
	TRIG :	BOOL;

	func_block : FT_TN8;
  END_VAR
	func_block.IN  :=IN ;
	func_block.T  :=T ;
	func_block();
	OUT := func_block.OUT;
	TRIG := func_block.TRIG;
END_PROGRAM

CONFIGURATION Config0

	VAR_GLOBAL
		PLC_TICKS_PER_SEC :	INT;
		PLC_SYS_TICK_CNT :	DINT;
	END_VAR

	RESOURCE Res0 ON PLC
		TASK task0(INTERVAL := T#20ms,PRIORITY := 0);
		PROGRAM instance0 WITH task0 : program0;
	END_RESOURCE

END_CONFIGURATION

(* ---- 546-FT_TN16.ST ---- *)
TYPE
  	oscat_arr_0_15               : ARRAY [0..15]    OF REAL;
END_TYPE

FUNCTION_BLOCK T_PLC_MS_Block
	VAR_OUTPUT
		T_PLC_MS :	UDINT;
	END_VAR

	VAR_EXTERNAL
		PLC_TICKS_PER_SEC :	INT;
		PLC_SYS_TICK_CNT :	DINT;
	END_VAR

	VAR
		debug :	BOOL;(*Debug-Mode ON / OFF*)
		N :	INT;(*Debug-Faktor*)
		Offset :	UDINT;(*Debug-Offset*)
		temp :	DWORD := DWORD#1;(*Debug-Offset*)
		mode :	BOOL;(*modus*)
		faktor :	UDINT;(*Systemtakt-Faktor*)
		init :	BOOL;
		v_plc_ticks_per_sec :	UDINT;
		base :	UDINT := UDINT#1000;
	END_VAR

	IF init = FALSE THEN
		v_plc_ticks_per_sec := INT_TO_UDINT(PLC_TICKS_PER_SEC);
		IF v_plc_ticks_per_sec = UDINT#1024 THEN
			faktor := UDINT#1;
			mode := FALSE;
		ELSIF v_plc_ticks_per_sec > UDINT#0 THEN
			IF v_plc_ticks_per_sec <= base THEN
				faktor := base / v_plc_ticks_per_sec;
				mode := FALSE;
			ELSE
				faktor := v_plc_ticks_per_sec / base;
				mode := TRUE;
			END_IF;
		ELSE
			faktor := UDINT#1;
		END_IF;
		init := TRUE;
	END_IF;

	IF mode THEN
		T_PLC_MS := DINT_TO_UDINT(PLC_SYS_TICK_CNT) / faktor;
	ELSE
		T_PLC_MS := DINT_TO_UDINT(PLC_SYS_TICK_CNT) * faktor;
	END_IF;

	IF debug THEN
		T_PLC_MS := (DWORD_TO_UDINT(SHL(UDINT_TO_DWORD(T_PLC_MS),N) OR SHL(temp,N)) - UDINT#1) + Offset;
	END_IF;
END_FUNCTION_BLOCK

FUNCTION_BLOCK FT_TN16
	VAR_INPUT
		IN :	REAL;
		T :	TIME;
	END_VAR

	VAR_OUTPUT
		OUT :	REAL;
		TRIG :	BOOL;
	END_VAR

	VAR
		length :	INT := 16;
		X :	oscat_arr_0_15;
		cnt :	INT;
		last :	TIME;
		tx :	TIME;
		init :	BOOL;
		T_PLC_MS :	T_PLC_MS_Block;
	END_VAR

	T_PLC_MS();
	tx:= UDINT_TO_TIME(T_PLC_MS.T_PLC_MS);

	trig := FALSE;
	IF NOT init THEN
		x[cnt] := in;
		init := TRUE;
		last := tx;
	ELSIF tx - last >= T / length THEN
		IF cnt = length - 1 THEN cnt := 0; ELSE cnt := cnt + 1; END_IF;
		Out := X[cnt];
		x[cnt] := in;
		last := tx;
		Trig := TRUE;
	END_IF;

END_FUNCTION_BLOCK

PROGRAM program0
  VAR
	IN :	REAL;
	T :	TIME;

	OUT :	REAL;
	TRIG :	BOOL;

	func_block : FT_TN16;
  END_VAR
	func_block.IN  :=IN ;
	func_block.T  :=T ;
	func_block();
	OUT := func_block.OUT;
	TRIG := func_block.TRIG;
END_PROGRAM

CONFIGURATION Config0

	VAR_GLOBAL
		PLC_TICKS_PER_SEC :	INT;
		PLC_SYS_TICK_CNT :	DINT;
	END_VAR

	RESOURCE Res0 ON PLC
		TASK task0(INTERVAL := T#20ms,PRIORITY := 0);
		PROGRAM instance0 WITH task0 : program0;
	END_RESOURCE

END_CONFIGURATION

(* ---- 547-FT_TN64.ST ---- *)
TYPE
	oscat_FT_TN64_array         : ARRAY [0..63]   OF REAL;
END_TYPE

FUNCTION_BLOCK T_PLC_MS_Block
	VAR_OUTPUT
		T_PLC_MS :	UDINT;
	END_VAR

	VAR_EXTERNAL
		PLC_TICKS_PER_SEC :	INT;
		PLC_SYS_TICK_CNT :	DINT;
	END_VAR

	VAR
		debug :	BOOL;(*Debug-Mode ON / OFF*)
		N :	INT;(*Debug-Faktor*)
		Offset :	UDINT;(*Debug-Offset*)
		temp :	DWORD := DWORD#1;(*Debug-Offset*)
		mode :	BOOL;(*modus*)
		faktor :	UDINT;(*Systemtakt-Faktor*)
		init :	BOOL;
		v_plc_ticks_per_sec :	UDINT;
		base :	UDINT := UDINT#1000;
	END_VAR

	IF init = FALSE THEN
		v_plc_ticks_per_sec := INT_TO_UDINT(PLC_TICKS_PER_SEC);
		IF v_plc_ticks_per_sec = UDINT#1024 THEN
			faktor := UDINT#1;
			mode := FALSE;
		ELSIF v_plc_ticks_per_sec > UDINT#0 THEN
			IF v_plc_ticks_per_sec <= base THEN
				faktor := base / v_plc_ticks_per_sec;
				mode := FALSE;
			ELSE
				faktor := v_plc_ticks_per_sec / base;
				mode := TRUE;
			END_IF;
		ELSE
			faktor := UDINT#1;
		END_IF;
		init := TRUE;
	END_IF;

	IF mode THEN
		T_PLC_MS := DINT_TO_UDINT(PLC_SYS_TICK_CNT) / faktor;
	ELSE
		T_PLC_MS := DINT_TO_UDINT(PLC_SYS_TICK_CNT) * faktor;
	END_IF;

	IF debug THEN
		T_PLC_MS := (DWORD_TO_UDINT(SHL(UDINT_TO_DWORD(T_PLC_MS),N) OR SHL(temp,N)) - UDINT#1) + Offset;
	END_IF;
END_FUNCTION_BLOCK

FUNCTION_BLOCK FT_TN64

	VAR_INPUT
		IN :	REAL;
		_T :	TIME;
	END_VAR

	VAR_OUTPUT
		OUT :	REAL;
		TRIG :	BOOL;
	END_VAR

	VAR
		length :	INT := 64;
		X :	oscat_FT_TN64_array;
		cnt :	INT;
		last :	TIME;
		tx :	TIME;
		init :	BOOL;
		T_PLC_MS :	T_PLC_MS_Block;
	END_VAR

	T_PLC_MS();
	tx:= UDINT_TO_TIME(T_PLC_MS.T_PLC_MS);

	trig := FALSE;
	IF NOT init THEN
		x[cnt] := in;
		init := TRUE;
		last := tx;
	ELSIF tx - last >= (_T / length) THEN
		IF cnt = length - 1 THEN cnt := 0; ELSE cnt := cnt + 1; END_IF;
		Out := X[cnt];
		x[cnt] := in;
		last := tx;
		trig := TRUE;
	END_IF;

END_FUNCTION_BLOCK

PROGRAM program0
  VAR
	IN :	REAL;
	_T :	TIME;

	OUT :	REAL;
	TRIG :	BOOL;

	func_block : FT_TN64;
  END_VAR
	func_block.IN  :=IN ;
	func_block._T  :=_T ;
	func_block();
	OUT := func_block.OUT;
	TRIG := func_block.TRIG;
END_PROGRAM

CONFIGURATION Config0

	VAR_GLOBAL
		PLC_TICKS_PER_SEC :	INT;
		PLC_SYS_TICK_CNT :	DINT;
	END_VAR

	RESOURCE Res0 ON PLC
		TASK task0(INTERVAL := T#20ms,PRIORITY := 0);
		PROGRAM instance0 WITH task0 : program0;
	END_RESOURCE

END_CONFIGURATION

(* ---- 548-RTC_MS.ST ---- *)
FUNCTION_BLOCK T_PLC_MS_Block
	VAR_OUTPUT
		T_PLC_MS :	UDINT;
	END_VAR

	VAR_EXTERNAL
		PLC_TICKS_PER_SEC :	INT;
		PLC_SYS_TICK_CNT :	DINT;
	END_VAR

	VAR
		debug :	BOOL;(*Debug-Mode ON / OFF*)
		N :	INT;(*Debug-Faktor*)
		Offset :	UDINT;(*Debug-Offset*)
		temp :	DWORD := DWORD#1;(*Debug-Offset*)
		mode :	BOOL;(*modus*)
		faktor :	UDINT;(*Systemtakt-Faktor*)
		init :	BOOL;
		v_plc_ticks_per_sec :	UDINT;
		base :	UDINT := UDINT#1000;
	END_VAR

	IF init = FALSE THEN
		v_plc_ticks_per_sec := INT_TO_UDINT(PLC_TICKS_PER_SEC);
		IF v_plc_ticks_per_sec = UDINT#1024 THEN
			faktor := UDINT#1;
			mode := FALSE;
		ELSIF v_plc_ticks_per_sec > UDINT#0 THEN
			IF v_plc_ticks_per_sec <= base THEN
				faktor := base / v_plc_ticks_per_sec;
				mode := FALSE;
			ELSE
				faktor := v_plc_ticks_per_sec / base;
				mode := TRUE;
			END_IF;
		ELSE
			faktor := UDINT#1;
		END_IF;
		init := TRUE;
	END_IF;

	IF mode THEN
		T_PLC_MS := DINT_TO_UDINT(PLC_SYS_TICK_CNT) / faktor;
	ELSE
		T_PLC_MS := DINT_TO_UDINT(PLC_SYS_TICK_CNT) * faktor;
	END_IF;

	IF debug THEN
		T_PLC_MS := (DWORD_TO_UDINT(SHL(UDINT_TO_DWORD(T_PLC_MS),N) OR SHL(temp,N)) - UDINT#1) + Offset;
	END_IF;
END_FUNCTION_BLOCK

FUNCTION_BLOCK RTC_MS_Block

	VAR_INPUT
		SET :	BOOL;
		SDT :	UDINT;
		SMS :	INT;
	END_VAR

	VAR_OUTPUT
		XDT :	UDINT;
		XMS :	INT;
	END_VAR

	VAR
		init :	BOOL;
		last :	UDINT;
		tx :	UDINT;
		T_PLC_MS :	T_PLC_MS_Block;
	END_VAR

	T_PLC_MS();
	tx:= T_PLC_MS.T_PLC_MS;

	IF set OR NOT init THEN
		(* clock needs to be set when set is true or after power up *)
		init := TRUE;
		xdt := SDT;
		XMS := SMS;
	ELSE
		XMS := XMS + UDINT_TO_INT(tx - last);
		(* check if one second has expired *)
		IF XMS > 999 THEN
			XDT := XDT + UDINT#1; (* add one second *)
			XMS := XMS - 1000;
		END_IF;
	END_IF;
	last := tx;

END_FUNCTION_BLOCK

PROGRAM program0

	VAR
		SET :	BOOL;
		SDT :	UDINT;
		SMS :	INT;
		XDT :	UDINT;
		XMS :	INT;
		func_block : RTC_MS_Block;
  	END_VAR
	func_block.SET  :=	SET;
	func_block.SDT  :=	SDT;
	func_block.SMS  :=	SMS;
	func_block();
	XDT := func_block.XDT;
	XMS := func_block.XMS;

END_PROGRAM

CONFIGURATION Config0

	VAR_GLOBAL
		PLC_TICKS_PER_SEC :	INT;
		PLC_SYS_TICK_CNT :	DINT;
	END_VAR

	RESOURCE Res0 ON PLC
		TASK task0(INTERVAL := T#20ms,PRIORITY := 0);
		PROGRAM instance0 WITH task0 : program0;
	END_RESOURCE

END_CONFIGURATION

(* ---- 550-CACOS.ST ---- *)
TYPE oscat_complex :
  STRUCT
	re : REAL;
	im : REAL;
  END_STRUCT;
END_TYPE

FUNCTION ATAN2:REAL
	VAR_INPUT
		X :	REAL;
		Y :	REAL;
	END_VAR

	IF X > 0.0 THEN
		ATAN2 := ATAN(Y/X);
	ELSIF X < 0.0 THEN
		IF Y >= 0.0 THEN
			ATAN2 := ATAN(Y/X) + 3.14159265358979323846264338327950288;
		ELSE
			ATAN2 := ATAN(Y/X) - 3.14159265358979323846264338327950288;
		END_IF;
	ELSIF Y > 0.0 THEN
		ATAN2 := 1.5707963267948965580;
	ELSIF Y < 0.0 THEN
		ATAN2 := -1.5707963267948965580;
	ELSE
		ATAN2 := 0.0;
	END_IF;

END_FUNCTION

FUNCTION HYPOT:REAL
	VAR_INPUT
		X :	REAL;
		Y :	REAL;
	END_VAR

	HYPOT := SQRT(x*x + y*y);
END_FUNCTION

FUNCTION_BLOCK CLOG_Block

	VAR_INPUT
		X :	oscat_complex;
	END_VAR

	VAR_OUTPUT
		CLOG :	oscat_complex;
	END_VAR

	CLOG.re := LN(HYPOT(X.re, X.im));
	CLOG.im := ATAN2(X.im, X.re);

END_FUNCTION_BLOCK

FUNCTION SGN : INT
  VAR_INPUT
    x : REAL;
  END_VAR

  IF X > 0.0 THEN
  	sgn := 1;
  ELSIF X < 0.0 THEN
  	sgn := -1;
  ELSE
  	sgn := 0;
  END_IF;
END_FUNCTION

FUNCTION_BLOCK CSQRT_Block
	VAR_INPUT
		X :	oscat_complex;
	END_VAR

	VAR_OUTPUT
		CSQRT :	oscat_complex;
	END_VAR

	VAR
		temp :	REAL;
	END_VAR

	temp := HYPOT(x.re, x.im);
	CSQRT.re :=  SQRT(0.5 * (temp + x.re));
	CSQRT.im :=  INT_TO_REAL(sgn(x.im)) * SQRT(0.5 * (temp - x.re));

END_FUNCTION_BLOCK

FUNCTION_BLOCK CACOSH_Block
	VAR_INPUT
		X :	oscat_complex;
	END_VAR

	VAR_OUTPUT
		CACOSH :	oscat_complex;
	END_VAR

	VAR
		Y :	oscat_complex;
		CLOG :	CLOG_Block;
		CSQRT :	CSQRT_Block;
	END_VAR

	y.re := (X.re - X.im)*(X.re + X.im) - 1.0;
	y.im := 2.0 * X.re * X.im;
	CSQRT(X:=y);
	y    := CSQRT.CSQRT;
	y.re := y.re + x.re;
	y.im := y.im + x.im;
	CLOG(X:=y);
	CACOSH  := CLOG.CLOG;
END_FUNCTION_BLOCK

FUNCTION_BLOCK CACOS_Block
	VAR_INPUT
		X :	oscat_complex;
	END_VAR

	VAR_OUTPUT
		CACOS :	oscat_complex;
	END_VAR

	VAR
		Y :	oscat_complex;
		CACOSH :	CACOSH_Block;
	END_VAR

	CACOSH(X:=x);
	y := CACOSH.CACOSH;
	CACOS.re := y.im;
	CACOS.im := -y.re;
END_FUNCTION_BLOCK

PROGRAM program0
  VAR
    LocalVar0 : oscat_complex;
	LocalOUT  : oscat_complex;
	func_block : CACOS_Block;
  END_VAR
	func_block.X  := LocalVar0;
	func_block();
	LocalOUT := func_block.CACOS;
END_PROGRAM

CONFIGURATION Config0
  RESOURCE Res0 ON PLC
    TASK task0(INTERVAL := T#20ms,PRIORITY := 0);
    PROGRAM instance0 WITH task0 : program0;
  END_RESOURCE
END_CONFIGURATION

(* ---- 551-NET_VAR_X8.ST ---- *)
FUNCTION_BLOCK NET_VAR_X8

	VAR_INPUT
		IN_REAL1 :	REAL;
		IN_REAL2 :	REAL;
		IN_DINT1 :	DINT;
		IN_DINT2 :	DINT;
		IN_UDINT1 :	UDINT;
		IN_UDINT2 :	UDINT;
		IN_DWORD1 :	DWORD;
		IN_DWORD2 :	DWORD;
	END_VAR

	VAR_OUTPUT
		OUT_REAL1 :	REAL;
		OUT_REAL2 :	REAL;
		OUT_DINT1 :	DINT;
		OUT_DINT2 :	DINT;
		OUT_UDINT1 :	UDINT;
		OUT_UDINT2 :	UDINT;
		OUT_DWORD1 :	DWORD;
		OUT_DWORD2 :	DWORD;
		ID :	BYTE;
	END_VAR

	VAR_IN_OUT
		X :	oscat_NET_VAR_DATA;
	END_VAR

	VAR
		init :	BOOL;
		i :	INT;
		i2 :	INT;
		index :	INT;
		index2 :	INT;
		REAL_TO_DW :	REAL_TO_DW;
		DW_TO_REAL :	DW_TO_REAL;
		ra :	oscat_nv_dw;
	END_VAR

	IF NOT init THEN
		init := TRUE;
		X.ID_MAX := X.ID_MAX + USINT#1;
		ID := USINT_TO_BYTE(X.ID_MAX);
	END_IF;

	IF X.STATE > BYTE#0 AND X.ERROR_ID = BYTE#0 THEN
		index := X.index;
		IF INT_TO_UINT(index + 34) > X.BUF_SIZE THEN
			X.ERROR_ID := ID;
		ELSE
			IF X.STATE = BYTE#1 THEN
				REAL_TO_DW(X:=IN_REAL1);
				ra[1] := REAL_TO_DW.REAL_TO_DW;
				REAL_TO_DW(X:=IN_REAL2);
				ra[2] := REAL_TO_DW.REAL_TO_DW;
				ra[3] := DINT_TO_DWORD(IN_DINT1);
				ra[4] := DINT_TO_DWORD(IN_DINT2);
				ra[5] := UDINT_TO_DWORD(IN_UDINT1);
				ra[6] := UDINT_TO_DWORD(IN_UDINT2);
				ra[7] := IN_DWORD1;
				ra[8] := IN_DWORD2;
				X.S_BUF.BUFFER[index] := ID;
				index := index + 1;
				X.S_BUF.BUFFER[index] := BYTE#21;
				index := index + 1;
				FOR i2 := 1 TO 8 DO;
					FOR i := 1 TO 4 DO;
						X.S_BUF.BUFFER[index] := DWORD_TO_BYTE(ra[i2]);
						ra[i2] := ROR(ra[i2],8);
						index := index + 1;
					END_FOR;
				END_FOR;

			ELSIF X.STATE = BYTE#2 THEN
				index2 := index + 1;
				IF X.R_BUF.BUFFER[index] <> ID OR X.R_BUF.BUFFER[index2] <> BYTE#21 THEN
					X.ERROR_ID := ID;
				ELSE
					index := index + 2;
					FOR i2 := 1 TO 8 DO;
						ra[i2] := DWORD#0;
						FOR i := 1 TO 4 DO;
							ra[i2] := ra[i2] OR BYTE_TO_DWORD(X.R_BUF.BUFFER[index]);
							ra[i2] := ROR(ra[i2],8);
							index := index + 1;
						END_FOR;
					END_FOR;
					DW_TO_REAL(X:=ra[1]);
					OUT_REAL1 := DW_TO_REAL.DW_TO_REAL;
					DW_TO_REAL(X:=ra[2]);
					OUT_REAL2 := DW_TO_REAL.DW_TO_REAL;
					OUT_DINT1 := DWORD_TO_DINT(ra[3]);
					OUT_DINT2 := DWORD_TO_DINT(ra[4]);
					OUT_UDINT1 := DWORD_TO_UDINT(ra[5]);
					OUT_UDINT2 := DWORD_TO_UDINT(ra[6]);
					OUT_DWORD1 := ra[7];
					OUT_DWORD2 := ra[8];
				END_IF;
			END_IF;
			X.index := index;
		END_IF;
	END_IF;

END_FUNCTION_BLOCK

(* ---- 552-CASIN.ST ---- *)
TYPE oscat_complex :
  STRUCT
	re : REAL;
	im : REAL;
  END_STRUCT;
END_TYPE

FUNCTION ATAN2:REAL
	VAR_INPUT
		X :	REAL;
		Y :	REAL;
	END_VAR

	IF X > 0.0 THEN
		ATAN2 := ATAN(Y/X);
	ELSIF X < 0.0 THEN
		IF Y >= 0.0 THEN
			ATAN2 := ATAN(Y/X) + 3.14159265358979323846264338327950288;
		ELSE
			ATAN2 := ATAN(Y/X) - 3.14159265358979323846264338327950288;
		END_IF;
	ELSIF Y > 0.0 THEN
		ATAN2 := 1.5707963267948965580;
	ELSIF Y < 0.0 THEN
		ATAN2 := -1.5707963267948965580;
	ELSE
		ATAN2 := 0.0;
	END_IF;

END_FUNCTION

FUNCTION HYPOT:REAL
	VAR_INPUT
		X :	REAL;
		Y :	REAL;
	END_VAR

	HYPOT := SQRT(x*x + y*y);
END_FUNCTION

FUNCTION_BLOCK CLOG_Block

	VAR_INPUT
		X :	oscat_complex;
	END_VAR

	VAR_OUTPUT
		CLOG :	oscat_complex;
	END_VAR

	CLOG.re := LN(HYPOT(X.re, X.im));
	CLOG.im := ATAN2(X.im, X.re);

END_FUNCTION_BLOCK

FUNCTION SGN : INT
  VAR_INPUT
    x : REAL;
  END_VAR

  IF X > 0.0 THEN
  	sgn := 1;
  ELSIF X < 0.0 THEN
  	sgn := -1;
  ELSE
  	sgn := 0;
  END_IF;
END_FUNCTION

FUNCTION_BLOCK CSQRT_Block
	VAR_INPUT
		X :	oscat_complex;
	END_VAR

	VAR_OUTPUT
		CSQRT :	oscat_complex;
	END_VAR

	VAR
		temp :	REAL;
	END_VAR

	temp := HYPOT(x.re, x.im);
	CSQRT.re :=  SQRT(0.5 * (temp + x.re));
	CSQRT.im :=  INT_TO_REAL(sgn(x.im)) * SQRT(0.5 * (temp - x.re));

END_FUNCTION_BLOCK

FUNCTION_BLOCK CASINH_Block
	VAR_INPUT
		X :	oscat_complex;
	END_VAR

	VAR_OUTPUT
		CASINH :	oscat_complex;
	END_VAR

	VAR
		Y :	oscat_complex;
		CLOG :	CLOG_Block;
		CSQRT :	CSQRT_Block;
	END_VAR

	y.re := (X.re - X.im)*(X.re + X.im) + 1.0;
	y.im := 2.0 * X.re * X.im;
	CSQRT(X:=y);
	y    := CSQRT.CSQRT;
	y.re := y.re + x.re;
	y.im := y.im + x.im;
	CLOG(X:=y);
	CASINH  := CLOG.CLOG;
END_FUNCTION_BLOCK

FUNCTION_BLOCK CASIN_Block
	VAR_INPUT
		X :	oscat_complex;
	END_VAR

	VAR_OUTPUT
		CASIN :	oscat_complex;
	END_VAR

	VAR
		Y :	oscat_complex;
		CASINH :	CASINH_Block;
	END_VAR

	y.re := -x.im;
	y.im := x.re;
	CASINH(X:=y);
	y := CASINH.CASINH;
	CASIN.re := y.im;
	CASIN.im := -y.re;
END_FUNCTION_BLOCK

PROGRAM program0
  VAR
    LocalVar0 : oscat_complex;
	LocalOUT  : oscat_complex;
	func_block : CASIN_Block;
  END_VAR
	func_block.X  := LocalVar0;
	func_block();
	LocalOUT := func_block.CASIN;
END_PROGRAM

CONFIGURATION Config0
  RESOURCE Res0 ON PLC
    TASK task0(INTERVAL := T#20ms,PRIORITY := 0);
    PROGRAM instance0 WITH task0 : program0;
  END_RESOURCE
END_CONFIGURATION

(* ---- 553-STRING_TO_TIME.ST ---- *)
FUNCTION_BLOCK UPPERCASE_Block

	VAR_INPUT
		STR :	STRING;
	END_VAR

	VAR_OUTPUT
		UPPERCASE :	STRING;
	END_VAR

	VAR
		char :	BYTE;
		char2 :	BYTE;
		pos :	INT;
		l :	INT;
		str_temp :	STRING;
	END_VAR

	UPPERCASE := str;
	l := LEN(str);
	FOR pos := 1 TO l DO
		char := INT_TO_BYTE(GET_CHAR(str,pos));
		char2 := TO_UPPER(char);
		IF char <> char2 THEN
			str_temp := UPPERCASE;
			UPPERCASE := REPLACE(str_temp,BYTE_TO_STRING(char2,'%c'),1,pos);
		END_IF;
	END_FOR;

END_FUNCTION_BLOCK

FUNCTION_BLOCK _STRING_TO_TIME
  VAR_INPUT
    _TIME :	STRING;
  END_VAR

  VAR_OUTPUT
    STRING_TO_TIME_O :	TIME;
  END_VAR

  VAR
    pos1 :	INT;
    pos2 :	INT;
    tmp :	STRING;
    tmp2 :	STRING;
    UPPERCASE :	UPPERCASE_Block;
    FINDB_NONUM :	FINDB_NONUM;
    FINDB_NUM :	FINDB_NUM;
    faktor :	UDINT;
    IS_ALNUM :	IS_ALNUM;
  END_VAR

  UPPERCASE(str:=_TIME);
  tmp:=UPPERCASE.UPPERCASE;

  STRING_TO_TIME_O := T#0s;

  WHILE (TRUE) DO
    FAKTOR := UDINT#0;

    FINDB_NONUM(str:=tmp);
    pos2:=FINDB_NONUM.findB_nonum;

    FINDB_NUM(str:=tmp);
    pos1:=FINDB_NUM.findB_num;

    (* bezeichner gefunden *)
    IF POS1>0 AND (POS2>POS1) THEN

      tmp2 := RIGHT(tmp,POS2-POS1);
      tmp := LEFT(tmp,pos1);

      IF EQ_STRING(tmp2,'MS') THEN
      FAKTOR := UDINT#1;
      ELSIF EQ_STRING(tmp2,'S') THEN
      FAKTOR := UDINT#1000;
      ELSIF EQ_STRING(tmp2,'M') THEN
      FAKTOR := UDINT#60000;
      ELSIF EQ_STRING(tmp2,'H') THEN
      FAKTOR := UDINT#3600000;
      ELSIF EQ_STRING(tmp2,'D') THEN
      FAKTOR := UDINT#864000000;
      END_IF;
    ELSE
      EXIT;
    END_IF;

    IF FAKTOR > UDINT#0 THEN

      FINDB_NONUM(str:=tmp);
      pos1:=FINDB_NONUM.findB_nonum;
      IF pos1>0 THEN
        tmp2 := RIGHT(tmp,LEN(tmp)-pos1);
        tmp := LEFT(tmp,pos1);
        IS_ALNUM(str:=tmp2);
        IF IS_ALNUM.IS_ALNUM THEN
          STRING_TO_TIME_O := STRING_TO_TIME_O + UDINT_TO_TIME(faktor * STRING_TO_UDINT(tmp2));
        END_IF;
      ELSE
      EXIT;
      END_IF;
    END_IF;
  END_WHILE;
END_FUNCTION_BLOCK

PROGRAM program0
	VAR
    LocalVar1 : STRING;
		LocalOUT  : TIME;
		func_block : _INSERT80;
  	END_VAR
	func_block._TIME := LocalVar1;
	func_block();
	LocalOUT := func_block.STRING_TO_TIME_O;
END_PROGRAM

CONFIGURATION Config0
  	RESOURCE Res0 ON PLC
    	TASK task0(INTERVAL := T#20ms,PRIORITY := 0);
    	PROGRAM instance0 WITH task0 : program0;
  	END_RESOURCE
END_CONFIGURATION

(* ---- 554-BASE64_DECODE_STR.ST ---- *)
TYPE
  oscat_aB0_47	: ARRAY [0..47]	OF BYTE;
  oscat_aB0_63	: ARRAY [0..63]	OF BYTE;
END_TYPE

FUNCTION_BLOCK BASE64_DECODE_STREAM
	VAR_IN_OUT
		BUF1 :	oscat_aB0_63;
		BUF2 :	oscat_aB0_47;
	END_VAR

	VAR_INPUT
		SIZE1 :	INT;
	END_VAR

	VAR_OUTPUT
		SIZE2 :	INT;
	END_VAR

	VAR
		a :	INT;
		b :	WORD;
		o :	INT;
		off :	INT;
		i1 :	INT;
		i2 :	INT;
		c :	INT;
	END_VAR

	IF SIZE1 <= 0 THEN SIZE2 := 0; RETURN; END_IF;
	c := SIZE1 - 1;
	i2 := 0;
	a := 0;
	b := WORD#0;
	FOR i1 := 0 TO c DO
		o := BYTE_TO_INT(BUF1[i1]);
		IF o = 61  (* = *) THEN EXIT;
		ELSIF o > 96 (* a-z *) THEN off := 71;
		ELSIF o > 64 (* A-Z *) THEN off := 65;
		ELSIF o > 47 (* 0-9 *) THEN off := -4;
		ELSIF o = 43 (* + *) THEN off := -19;
		ELSIF o = 47 (* / *) THEN off := -16;
		END_IF;
		b := SHL(b,6) OR INT_TO_WORD(o - off);
		a := a + 6;
		IF a >= 8 THEN
			a := a - 8;
			BUF2[i2] := WORD_TO_BYTE(SHR(b,a));
			i2 := i2 + 1;
			b := b AND NOT SHL(WORD#16#FFFF,a);
		END_IF;
	END_FOR;
	SIZE2 := i2;
END_FUNCTION_BLOCK

FUNCTION_BLOCK BASE64_DECODE_STR
	VAR_INPUT
		RUN :	BOOL;
	END_VAR

	VAR_OUTPUT
		DONE :	BOOL;
	END_VAR

	VAR_IN_OUT
		STR1 :	STRING;
		STR2 :	STRING;
	END_VAR

	VAR
		BASE64_DECODE_STREAM :	BASE64_DECODE_STREAM;
		run_last :	BOOL;
		buf1 :	oscat_aB0_63;
		buf2 :	oscat_aB0_47;
		mode :	INT;
		size1 :	INT;
		size2 :	INT;
		end :	INT;
		pos :	INT;
		i1 :	INT;
		i2 :	INT;
		i3 :	INT;
		STRx :	STRING;
		BTS :	BUF_TO_STRING;
	END_VAR

	(*@KEY@: WORKSHEET
	NAME: BASE64_DECODE_STR
	IEC_LANGUAGE: ST
	*)

	CASE mode OF
	0:	IF RUN AND NOT run_last THEN
			DONE := FALSE;
			mode := 1;
			end := LEN(STR1);
			pos := 0;
			STR2 := '';
		END_IF;
	1:
		SIZE1 := MIN(48,end - pos);
		IF SIZE1 > 0 THEN

			i2 := SIZE1 - 1;
			i3 := pos + 1;
			FOR i1 := 0 TO i2 DO
				buf1[i1] := INT_TO_BYTE(GET_CHAR(STR1,i3));
				i3 := i3 + 1;
			END_FOR;

			BASE64_DECODE_STREAM(BUF1:=BUF1 ,BUF2:=BUF2 ,SIZE1:=SIZE1);
			buf1  :=BASE64_DECODE_STREAM.BUF1;
			buf2  :=BASE64_DECODE_STREAM.BUF2;
			SIZE2 :=BASE64_DECODE_STREAM.SIZE2;

			FOR i1 := 0 TO 1 DO
				BTS.REQ := i1 > 0;
				BTS.BUF_FORMAT := TRUE;
				BTS.BUF_OFFS := DINT#0;
				BTS.BUF_CNT := INT_TO_DINT(SIZE2);
				BTS.BUFFER := buf2;
				BTS.DST := STRx;
				BTS();
				buf2 := BTS.BUFFER;
				STRx := BTS.DST;
			END_FOR;
			STR2 := CONCAT(STR2,STRx);
		ELSE
			mode := 0;
			DONE := TRUE;
		END_IF;
		pos := pos + size1;
	END_CASE;

	run_last := RUN;

END_FUNCTION_BLOCK

(* ---- 555-ONTIME.ST ---- *)
FUNCTION_BLOCK T_PLC_MS_block
	VAR_OUTPUT
		T_PLC_MS :	UDINT;
	END_VAR

	VAR_EXTERNAL
		PLC_TICKS_PER_SEC :	INT;
		PLC_SYS_TICK_CNT :	DINT;
	END_VAR

	VAR
		debug :	BOOL;(*Debug-Mode ON / OFF*)
		N :	INT;(*Debug-Faktor*)
		Offset :	UDINT;(*Debug-Offset*)
		temp :	DWORD := DWORD#1;(*Debug-Offset*)
		mode :	BOOL;(*modus*)
		faktor :	UDINT;(*Systemtakt-Faktor*)
		init :	BOOL;
		v_plc_ticks_per_sec :	UDINT;
		base :	UDINT := UDINT#1000;
	END_VAR

	IF init = FALSE THEN
		v_plc_ticks_per_sec := INT_TO_UDINT(PLC_TICKS_PER_SEC);
		IF v_plc_ticks_per_sec = UDINT#1024 THEN
			faktor := UDINT#1;
			mode := FALSE;
		ELSIF v_plc_ticks_per_sec > UDINT#0 THEN
			IF v_plc_ticks_per_sec <= base THEN
				faktor := base / v_plc_ticks_per_sec;
				mode := FALSE;
			ELSE
				faktor := v_plc_ticks_per_sec / base;
				mode := TRUE;
			END_IF;
		ELSE
			faktor := UDINT#1;
		END_IF;
		init := TRUE;
	END_IF;

	IF mode THEN
		T_PLC_MS := DINT_TO_UDINT(PLC_SYS_TICK_CNT) / faktor;
	ELSE
		T_PLC_MS := DINT_TO_UDINT(PLC_SYS_TICK_CNT) * faktor;
	END_IF;

	IF debug THEN
		T_PLC_MS := (DWORD_TO_UDINT(SHL(UDINT_TO_DWORD(T_PLC_MS),N) OR SHL(temp,N)) - UDINT#1) + Offset;
	END_IF;

END_FUNCTION_BLOCK

FUNCTION_BLOCK ONTIME_Block

	VAR_INPUT
		IN :	BOOL;
		RST :	BOOL;
	END_VAR

	VAR_IN_OUT
		SECONDS :	UDINT;
		CYCLES :	UDINT;
	END_VAR

	VAR
		tx :	UDINT;
		last :	UDINT;
		edge :	BOOL;
		init :	BOOL;
		ms :	UDINT;
		T_PLC_MS :	T_PLC_MS_Block;
	END_VAR

	T_PLC_MS();
	tx:= T_PLC_MS.T_PLC_MS;

	IF NOT init THEN
		init := TRUE;
		last := tx;
		ms := UDINT#0;
	END_IF;
	IF RST THEN
		SECONDS := UDINT#0;
		CYCLES := UDINT#0;
		last := tx;
		ms := UDINT#0;
	ELSIF IN THEN
		(* add the current milliseconds *)
		ms := (tx - last) + ms;
		IF ms >= UDINT#1000 THEN
			seconds := seconds + UDINT#1;
			ms := ms - UDINT#1000;
		END_IF;
		cycles := cycles + BOOL_TO_UDINT(NOT edge);
	END_IF;
	last := tx;
	edge := in;

END_FUNCTION_BLOCK

PROGRAM program0
	VAR
		IN :	BOOL;
		RST :	BOOL;
		SECONDS :	UDINT;
		CYCLES :	UDINT;
		func_block : ONTIME_Block;
	END_VAR
	func_block.IN := IN;
	func_block.RST := RST;
	func_block();
	SECONDS  := func_block.SECONDS;
	CYCLES  := func_block.CYCLES;
END_PROGRAM

CONFIGURATION Config0
	VAR_GLOBAL
		PLC_TICKS_PER_SEC :	INT;
		PLC_SYS_TICK_CNT :	DINT;
	END_VAR
  	RESOURCE Res0 ON PLC
    	TASK task0(INTERVAL := T#20ms,PRIORITY := 0);
    	PROGRAM instance0 WITH task0 : program0;
  	END_RESOURCE
END_CONFIGURATION

(* ---- 556-PULSE_T.ST ---- *)
FUNCTION UDINT_TO_TIME2:TIME

	VAR_INPUT
		IN :	UDINT;
	END_VAR

	UDINT_TO_TIME2 := DINT_TO_TIME(UDINT_TO_DINT(IN));

END_FUNCTION

FUNCTION_BLOCK T_PLC_MS_block
	VAR_OUTPUT
		T_PLC_MS :	UDINT;
	END_VAR

	VAR_EXTERNAL
		PLC_TICKS_PER_SEC :	INT;
		PLC_SYS_TICK_CNT :	DINT;
	END_VAR

	VAR
		debug :	BOOL;(*Debug-Mode ON / OFF*)
		N :	INT;(*Debug-Faktor*)
		Offset :	UDINT;(*Debug-Offset*)
		temp :	DWORD := DWORD#1;(*Debug-Offset*)
		mode :	BOOL;(*modus*)
		faktor :	UDINT;(*Systemtakt-Faktor*)
		init :	BOOL;
		v_plc_ticks_per_sec :	UDINT;
		base :	UDINT := UDINT#1000;
	END_VAR

	IF init = FALSE THEN
		v_plc_ticks_per_sec := INT_TO_UDINT(PLC_TICKS_PER_SEC);
		IF v_plc_ticks_per_sec = UDINT#1024 THEN
			faktor := UDINT#1;
			mode := FALSE;
		ELSIF v_plc_ticks_per_sec > UDINT#0 THEN
			IF v_plc_ticks_per_sec <= base THEN
				faktor := base / v_plc_ticks_per_sec;
				mode := FALSE;
			ELSE
				faktor := v_plc_ticks_per_sec / base;
				mode := TRUE;
			END_IF;
		ELSE
			faktor := UDINT#1;
		END_IF;
		init := TRUE;
	END_IF;

	IF mode THEN
		T_PLC_MS := DINT_TO_UDINT(PLC_SYS_TICK_CNT) / faktor;
	ELSE
		T_PLC_MS := DINT_TO_UDINT(PLC_SYS_TICK_CNT) * faktor;
	END_IF;

	IF debug THEN
		T_PLC_MS := (DWORD_TO_UDINT(SHL(UDINT_TO_DWORD(T_PLC_MS),N) OR SHL(temp,N)) - UDINT#1) + Offset;
	END_IF;

END_FUNCTION_BLOCK

FUNCTION_BLOCK PULSE_T_Block

	VAR_INPUT
		IN :	BOOL;
		T1 :	TIME;
		T2 :	TIME;
		RST :	BOOL;
	END_VAR

	VAR_OUTPUT
		Q :	BOOL;
	END_VAR

	VAR
		init :	BOOL;
		last :	TIME;
		tx :	TIME;
		edge :	BOOL;
		T_PLC_MS :	T_PLC_MS_Block;
	END_VAR

	T_PLC_MS();
	tx:= UDINT_TO_TIME(T_PLC_MS.T_PLC_MS);

	IF NOT init THEN
		init := TRUE;
		last := tx;
	ELSIF RST THEN
		Q := FALSE;
	ELSIF IN AND NOT edge AND NOT Q THEN
		last := tx;
		Q := TRUE;
	ELSIF NOT IN AND edge AND ((tx - last) > T1) THEN
		Q := FALSE;
	ELSIF (tx - last) >= T2 THEN
		Q := FALSE;
	END_IF;

	edge := IN;

END_FUNCTION_BLOCK

PROGRAM program0
	VAR
		IN :	BOOL;
		T1 :	TIME;
		T2 :	TIME;
		RST :	BOOL;
		Q :	BOOL;

		func_block : PULSE_T_Block;
	END_VAR
	func_block.IN := IN;
	func_block.T1 := T1;
	func_block.T2 := T2 ;
	func_block.RST := RST ;

	func_block();
	Q  := func_block.Q;
END_PROGRAM

CONFIGURATION Config0
	VAR_GLOBAL
		PLC_TICKS_PER_SEC :	INT;
		PLC_SYS_TICK_CNT :	DINT;
	END_VAR
  	RESOURCE Res0 ON PLC
    	TASK task0(INTERVAL := T#20ms,PRIORITY := 0);
    	PROGRAM instance0 WITH task0 : program0;
  	END_RESOURCE
END_CONFIGURATION

(* ---- 557-FIX.ST ---- *)
FUNCTION _BYTE_TO_INT:INT
	VAR_INPUT
		IN :	BYTE;
	END_VAR

	_BYTE_TO_INT := USINT_TO_INT(BYTE_TO_USINT(IN));
END_FUNCTION

FUNCTION_BLOCK CHR_TO_STRING_Block
	VAR_INPUT
		C :	BYTE;
	END_VAR

	VAR_OUTPUT
		CHR_TO_STRING :	STRING;
	END_VAR

	CHR_TO_STRING := BYTE_TO_STRING(C);

END_FUNCTION_BLOCK

FUNCTION BIT_OF_DWORD : BOOL
  VAR_INPUT
    IN : DWORD;
    N : INT;
  END_VAR

  BIT_OF_DWORD := (SHR(in,N) AND 16#00000001) > 0;
  (* from OSCAT library; www.oscat.de  *)
END_FUNCTION

FUNCTION_BLOCK FILL_Block
	VAR_INPUT
		C :	BYTE;
		L :	INT;
	END_VAR

	VAR_OUTPUT
		FILL :	STRING;
	END_VAR

	VAR
		N :	BYTE;
		I :	INT;
		sx :	STRING;
		CHR_TO_STRING :	CHR_TO_STRING_Block;
		FILL_tmp :	STRING;
	END_VAR

	CHR_TO_STRING(C:=c);
	Sx:=CHR_TO_STRING.CHR_TO_STRING;
	(* create string *)
	N := INT_TO_BYTE(LIMIT(0,L,80));
	(* create a string of characters to be connected to str *)
	FILL := '';
	FOR i := 1 TO 8 DO
		FILL_tmp := FILL;
		FILL := CONCAT(FILL_tmp,FILL);
		IF BIT_OF_DWORD(BYTE_TO_DWORD(N),7) THEN FILL := CONCAT(FILL,Sx); END_IF;
		N := SHL(N,1);
	END_FOR;
END_FUNCTION_BLOCK

FUNCTION_BLOCK FIX_Block

	VAR_INPUT
		STR :	STRING;
		L :	INT;
		C :	BYTE;
		M :	INT;
	END_VAR

	VAR_OUTPUT
		FIX :	STRING;
	END_VAR

	VAR
		N :	INT;
		FILL :	FILL_Block;
	END_VAR

	N := LIMIT(0,L,255) - LEN(str);
	IF N <= 0 THEN
		(* truncate the string at length N *)
		IF M = 1 THEN
			FIX := RIGHT(str,L);
		ELSE
			FIX := LEFT(str,L);
		END_IF;
	ELSIF M = 1 THEN
		(* connect fill characters at the beginning *)
		FILL(C:=C,L:=N);
		FIX := CONCAT(FILL.FILL,str);
	ELSIF M = 2 THEN
		(* center str beween fill characters *)
		(* for an uneven number of fill characters, there is one more at the end *)
		FILL(C:=C,L:=_BYTE_TO_INT(SHR(INT_TO_BYTE(N+1),1)));
		FIX := CONCAT(str,FILL.FILL);
		FILL(C:=C,L:=_BYTE_TO_INT(SHR(INT_TO_BYTE(N),1)));
		FIX := CONCAT(FILL.FILL,FIX);
	ELSE
		(* connect fill characters at the end *)
		FILL(C:=C,L:=N);
		FIX := CONCAT(str,FILL.FILL);
	END_IF;

END_FUNCTION_BLOCK

PROGRAM program0
  VAR
	STR :	STRING;
	L   :	INT;
	C   :	BYTE;
	M   :	INT;

	FIX :	STRING;

	func_block : FIX_Block;
  END_VAR
	func_block.STR:=STR;
	func_block.L  :=L  ;
	func_block.C  :=C  ;
	func_block.M  :=M  ;
	func_block();
	FIX := func_block.FIX;
END_PROGRAM

CONFIGURATION Config0
  RESOURCE Res0 ON PLC
    TASK task0(INTERVAL := T#20ms,PRIORITY := 0);
    PROGRAM instance0 WITH task0 : program0;
  END_RESOURCE
END_CONFIGURATION

(* ---- 559-TP_1D.ST ---- *)
FUNCTION UDINT_TO_TIME2:TIME

	VAR_INPUT
		IN :	UDINT;
	END_VAR

	UDINT_TO_TIME2 := DINT_TO_TIME(UDINT_TO_DINT(IN));

END_FUNCTION

FUNCTION_BLOCK T_PLC_MS_block
	VAR_OUTPUT
		T_PLC_MS :	UDINT;
	END_VAR

	VAR_EXTERNAL
		PLC_TICKS_PER_SEC :	INT;
		PLC_SYS_TICK_CNT :	DINT;
	END_VAR

	VAR
		debug :	BOOL;(*Debug-Mode ON / OFF*)
		N :	INT;(*Debug-Faktor*)
		Offset :	UDINT;(*Debug-Offset*)
		temp :	DWORD := DWORD#1;(*Debug-Offset*)
		mode :	BOOL;(*modus*)
		faktor :	UDINT;(*Systemtakt-Faktor*)
		init :	BOOL;
		v_plc_ticks_per_sec :	UDINT;
		base :	UDINT := UDINT#1000;
	END_VAR

	IF init = FALSE THEN
		v_plc_ticks_per_sec := INT_TO_UDINT(PLC_TICKS_PER_SEC);
		IF v_plc_ticks_per_sec = UDINT#1024 THEN
			faktor := UDINT#1;
			mode := FALSE;
		ELSIF v_plc_ticks_per_sec > UDINT#0 THEN
			IF v_plc_ticks_per_sec <= base THEN
				faktor := base / v_plc_ticks_per_sec;
				mode := FALSE;
			ELSE
				faktor := v_plc_ticks_per_sec / base;
				mode := TRUE;
			END_IF;
		ELSE
			faktor := UDINT#1;
		END_IF;
		init := TRUE;
	END_IF;

	IF mode THEN
		T_PLC_MS := DINT_TO_UDINT(PLC_SYS_TICK_CNT) / faktor;
	ELSE
		T_PLC_MS := DINT_TO_UDINT(PLC_SYS_TICK_CNT) * faktor;
	END_IF;

	IF debug THEN
		T_PLC_MS := (DWORD_TO_UDINT(SHL(UDINT_TO_DWORD(T_PLC_MS),N) OR SHL(temp,N)) - UDINT#1) + Offset;
	END_IF;

END_FUNCTION_BLOCK

FUNCTION_BLOCK TP_1D
	VAR_INPUT
		IN :	BOOL;
		PT1 :	TIME;
		PTD :	TIME;
		RST :	BOOL;
	END_VAR

	VAR_OUTPUT
		Q :	BOOL;
		W :	BOOL;
	END_VAR

	VAR
		tx :	TIME;
		start :	TIME;
		ix :	BOOL;
		T_PLC_MS :	T_PLC_MS_block;
	END_VAR

	T_PLC_MS();
	tx := UDINT_TO_TIME(T_PLC_MS.T_PLC_MS);

	IF RST THEN
		Q := FALSE;
		rst := FALSE;
		W := FALSE;
	ELSIF W THEN
		IF tx - start >= PTD THEN
			W := FALSE;
		END_IF;
	ELSIF IN AND NOT ix THEN
		Q := TRUE;
		start := tx;
		in := FALSE;
	ELSIF tx - start >= PT1 THEN
		Q := FALSE;
		W := TRUE;
		start := tx;
	END_IF;

	ix := IN;

END_FUNCTION_BLOCK

PROGRAM program0
  VAR
	IN :	BOOL;
	PT1 :	TIME;
	PTD :	TIME;
	RST :	BOOL;
	Q :	BOOL;
	W :	BOOL;
	func_block : TP_1D;
  END_VAR
	func_block.IN  :=IN;
	func_block.PT1  :=PT1;
	func_block.PTD  :=PTD;
	func_block.RST  :=RST;
	func_block();
	Q := func_block.Q;
	W := func_block.W;
END_PROGRAM

CONFIGURATION Config0
	VAR_GLOBAL
		PLC_TICKS_PER_SEC :	INT;
		PLC_SYS_TICK_CNT :	DINT;
	END_VAR
	RESOURCE Res0 ON PLC
		TASK task0(INTERVAL := T#20ms,PRIORITY := 0);
		PROGRAM instance0 WITH task0 : program0;
	END_RESOURCE
END_CONFIGURATION

(* ---- 560-CLK_PULSE.ST ---- *)
FUNCTION_BLOCK T_PLC_MS_block
	VAR_OUTPUT
		T_PLC_MS :	UDINT;
	END_VAR

	VAR_EXTERNAL
		PLC_TICKS_PER_SEC :	INT;
		PLC_SYS_TICK_CNT :	DINT;
	END_VAR

	VAR
		debug :	BOOL;(*Debug-Mode ON / OFF*)
		N :	INT;(*Debug-Faktor*)
		Offset :	UDINT;(*Debug-Offset*)
		temp :	DWORD := DWORD#1;(*Debug-Offset*)
		mode :	BOOL;(*modus*)
		faktor :	UDINT;(*Systemtakt-Faktor*)
		init :	BOOL;
		v_plc_ticks_per_sec :	UDINT;
		base :	UDINT := UDINT#1000;
	END_VAR

	IF init = FALSE THEN
		v_plc_ticks_per_sec := INT_TO_UDINT(PLC_TICKS_PER_SEC);
		IF v_plc_ticks_per_sec = UDINT#1024 THEN
			faktor := UDINT#1;
			mode := FALSE;
		ELSIF v_plc_ticks_per_sec > UDINT#0 THEN
			IF v_plc_ticks_per_sec <= base THEN
				faktor := base / v_plc_ticks_per_sec;
				mode := FALSE;
			ELSE
				faktor := v_plc_ticks_per_sec / base;
				mode := TRUE;
			END_IF;
		ELSE
			faktor := UDINT#1;
		END_IF;
		init := TRUE;
	END_IF;

	IF mode THEN
		T_PLC_MS := DINT_TO_UDINT(PLC_SYS_TICK_CNT) / faktor;
	ELSE
		T_PLC_MS := DINT_TO_UDINT(PLC_SYS_TICK_CNT) * faktor;
	END_IF;

	IF debug THEN
		T_PLC_MS := (DWORD_TO_UDINT(SHL(UDINT_TO_DWORD(T_PLC_MS),N) OR SHL(temp,N)) - UDINT#1) + Offset;
	END_IF;

END_FUNCTION_BLOCK

FUNCTION TIME_TO_UDINT2:UDINT
	VAR_INPUT
		X :	TIME;
	END_VAR

	TIME_TO_UDINT2 := DINT_TO_UDINT(TIME_TO_DINT(X));
END_FUNCTION

FUNCTION_BLOCK CLK_PULSE
	VAR_INPUT
		PT :	TIME;
		N :	INT;
		RST :	BOOL;
	END_VAR

	VAR_OUTPUT
		Q :	BOOL;
		CNT :	INT;
		RUN :	BOOL;
	END_VAR

	VAR
		tx :	UDINT;
		tn :	UDINT;
		init :	BOOL;
		T_PLC_MS :	T_PLC_MS_block;
	END_VAR

	T_PLC_MS();
	tx:= T_PLC_MS.T_PLC_MS;
	Q := FALSE;				(* reset Q we generate pulses only for one cycle *)
	RUN := CNT < N;

	IF NOT init OR RST THEN
		init := TRUE;
		CNT := 0;
		tn := tx - TIME_TO_UDINT2(PT);
		RUN := FALSE;
	ELSIF (cnt < N OR N = 0) AND tx - tn >= TIME_TO_UDINT2(PT) THEN		(* generate a pulse *)
		CNT := CNT + 1;
		Q := TRUE;
		tn := tn + TIME_TO_UDINT2(PT);
	END_IF;

END_FUNCTION_BLOCK

PROGRAM program0
  VAR
    LocalVar0 : TIME;
	LocalVar1 : INT;
	LocalVar2 : BOOL;

	Q :	BOOL;
	CNT :	INT;
	RUN :	BOOL;
	func_block : CLK_PULSE;
  END_VAR
	func_block.PT  := LocalVar0;
	func_block.N  := LocalVar1;
	func_block.RST  := LocalVar2;
	func_block();
	Q:= func_block.Q;
	CNT := func_block.CNT;
	RUN := func_block.RUN;

END_PROGRAM

CONFIGURATION Config0
	VAR_GLOBAL
		PLC_TICKS_PER_SEC :	INT;
		PLC_SYS_TICK_CNT :	DINT;
	END_VAR

  RESOURCE Res0 ON PLC
    TASK task0(INTERVAL := T#20ms,PRIORITY := 0);
    PROGRAM instance0 WITH task0 : program0;
  END_RESOURCE
END_CONFIGURATION

(* ---- 561-FT_PD.ST ---- *)
FUNCTION_BLOCK T_PLC_US_Block
	VAR_OUTPUT
		T_PLC_US :	UDINT;
	END_VAR

	VAR_EXTERNAL
		PLC_TICKS_PER_SEC :	INT;
		PLC_SYS_TICK_CNT :	DINT;
	END_VAR

	VAR
		debug :	BOOL;
		N :	INT;
		Offset :	UDINT;
		temp :	DWORD := DWORD#1;
		mode :	BOOL;
		faktor :	UDINT;
		init :	BOOL;
		v_plc_ticks_per_sec :	UDINT;
		base :	UDINT := UDINT#1000000;
	END_VAR

	IF init = FALSE THEN
		v_plc_ticks_per_sec := INT_TO_UDINT(PLC_TICKS_PER_SEC);
		IF v_plc_ticks_per_sec = UDINT#1024 THEN
			faktor := UDINT#1000;
			mode := FALSE;
		ELSIF v_plc_ticks_per_sec > UDINT#0 THEN
			IF v_plc_ticks_per_sec <= base THEN
				faktor := base / v_plc_ticks_per_sec;
				mode := FALSE;
			ELSE
				faktor := v_plc_ticks_per_sec / base;
				mode := TRUE;
			END_IF;
		ELSE
			faktor := UDINT#1;
		END_IF;
		init := TRUE;
	END_IF;

	IF mode THEN
		T_PLC_US := DINT_TO_UDINT(PLC_SYS_TICK_CNT) / faktor;
	ELSE
		T_PLC_US := DINT_TO_UDINT(PLC_SYS_TICK_CNT) * faktor;
	END_IF;

	IF debug THEN
		T_PLC_US := (DWORD_TO_UDINT(SHL(UDINT_TO_DWORD(T_PLC_US),N) OR SHL(temp,N)) - UDINT#1) + Offset;
	END_IF;
END_FUNCTION_BLOCK

FUNCTION_BLOCK FT_DERIV
	VAR_INPUT
		IN :	REAL;
		K :	REAL := 1.0;
		RUN :	BOOL := TRUE;
	END_VAR

	VAR_OUTPUT
		OUT :	REAL;
	END_VAR

	VAR
		old :	REAL;
		tx :	UDINT;
		last :	UDINT;
		init :	BOOL;
		tc :	REAL;
		T_PLC_US :	T_PLC_US_Block;
	END_VAR

	T_PLC_US();
	tx:= T_PLC_US.T_PLC_US;
	tc := UDINT_TO_REAL(tx - last);

	IF NOT init THEN
		init := TRUE;
		old := in;
	ELSIF run AND tc > 0.0 THEN
		out := (in - old) / tc * 1000000.0 * K;
		old := in;
	ELSE
		out := 0.0;
	END_IF;

	last := tx;

	T_PLC_US();
	tx:= T_PLC_US.T_PLC_US;

	IF NOT init THEN
		init := TRUE;
	ELSIF run AND tx - last > UDINT#0 THEN
		out := (in - old) / UDINT_TO_REAL(tx - last) * 1000000.0 * K;
	ELSE
		out := 0.0;
	END_IF;
	old := in;
	last := tx;
END_FUNCTION_BLOCK

FUNCTION_BLOCK FT_PD_Block

	VAR_INPUT
		IN :	REAL;
		KP :	REAL := 1.0;
		TV :	REAL := 1.0;
	END_VAR

	VAR_OUTPUT
		Y :	REAL;
	END_VAR

	VAR
		diff :	FT_DERIV;
	END_VAR

	diff(IN := IN, K := TV);

	Y := KP * (diff.out + IN);

END_FUNCTION_BLOCK

PROGRAM program0
	VAR
		IN :	REAL;
		KP :	REAL := 1.0;
		TV :	REAL := 1.0;
		Y :	REAL;
		func_block : FT_PD_Block;
	END_VAR
	func_block.IN :=IN;
	func_block.KP :=KP;
	func_block.TV :=TV;
	func_block();
	Y := func_block.Y;
END_PROGRAM

CONFIGURATION Config0

	VAR_GLOBAL
		PLC_TICKS_PER_SEC :	INT;
		PLC_SYS_TICK_CNT :	DINT;
	END_VAR

	RESOURCE Res0 ON PLC
		TASK task0(INTERVAL := T#20ms,PRIORITY := 0);
		PROGRAM instance0 WITH task0 : program0;
	END_RESOURCE

END_CONFIGURATION

(* ---- 562-FILTER_DW.ST ---- *)
FUNCTION_BLOCK T_PLC_MS_block
	VAR_OUTPUT
		T_PLC_MS :	UDINT;
	END_VAR

	VAR_EXTERNAL
		PLC_TICKS_PER_SEC :	INT;
		PLC_SYS_TICK_CNT :	DINT;
	END_VAR

	VAR
		debug :	BOOL;(*Debug-Mode ON / OFF*)
		N :	INT;(*Debug-Faktor*)
		Offset :	UDINT;(*Debug-Offset*)
		temp :	DWORD := DWORD#1;(*Debug-Offset*)
		mode :	BOOL;(*modus*)
		faktor :	UDINT;(*Systemtakt-Faktor*)
		init :	BOOL;
		v_plc_ticks_per_sec :	UDINT;
		base :	UDINT := UDINT#1000;
	END_VAR

	IF init = FALSE THEN
		v_plc_ticks_per_sec := INT_TO_UDINT(PLC_TICKS_PER_SEC);
		IF v_plc_ticks_per_sec = UDINT#1024 THEN
			faktor := UDINT#1;
			mode := FALSE;
		ELSIF v_plc_ticks_per_sec > UDINT#0 THEN
			IF v_plc_ticks_per_sec <= base THEN
				faktor := base / v_plc_ticks_per_sec;
				mode := FALSE;
			ELSE
				faktor := v_plc_ticks_per_sec / base;
				mode := TRUE;
			END_IF;
		ELSE
			faktor := UDINT#1;
		END_IF;
		init := TRUE;
	END_IF;

	IF mode THEN
		T_PLC_MS := DINT_TO_UDINT(PLC_SYS_TICK_CNT) / faktor;
	ELSE
		T_PLC_MS := DINT_TO_UDINT(PLC_SYS_TICK_CNT) * faktor;
	END_IF;

	IF debug THEN
		T_PLC_MS := (DWORD_TO_UDINT(SHL(UDINT_TO_DWORD(T_PLC_MS),N) OR SHL(temp,N)) - UDINT#1) + Offset;
	END_IF;

END_FUNCTION_BLOCK

FUNCTION _DWORD_TO_REAL:REAL
	VAR_INPUT
		IN :	DWORD;
	END_VAR

	_DWORD_TO_REAL := UDINT_TO_REAL(DWORD_TO_UDINT(IN));
END_FUNCTION

FUNCTION _REAL_TO_DWORD: DWORD

  VAR_INPUT
    X :	REAL;
  END_VAR

  IF REAL_TO_DWORD(0.5) = DWORD#1 THEN
    _REAL_TO_DWORD := REAL_TO_DWORD(x);
  ELSIF X > 0.0 THEN
    _REAL_TO_DWORD := REAL_TO_DWORD(x+0.5);
  ELSIF X < 0.0 THEN
    _REAL_TO_DWORD := REAL_TO_DWORD(x-0.5);
  ELSE
    _REAL_TO_DWORD := DWORD#0;
  END_IF;
END_FUNCTION

FUNCTION_BLOCK FILTER_DW

	VAR_INPUT
		X :	DWORD;
		T :	TIME;
	END_VAR

	VAR_OUTPUT
		Y :	DWORD;
	END_VAR

	VAR
		last :	UDINT;
		tx :	UDINT;
		init :	BOOL;
		Yi :	REAL;
		T_PLC_MS :	T_PLC_MS_block;
	END_VAR

	T_PLC_MS();
	tx:= T_PLC_MS.T_PLC_MS;

	IF NOT init OR T = t#0s THEN
		init := TRUE;
		Yi := _DWORD_TO_REAL(X);
	ELSE
		Yi := Yi + (_DWORD_TO_REAL(X) - _DWORD_TO_REAL(Y)) * UDINT_TO_REAL(tx - last) / TIME_TO_REAL(T);
	END_IF;
	last := tx;

	Y := _REAL_TO_DWORD(Yi);

END_FUNCTION_BLOCK

PROGRAM program0
  VAR
	X :	DWORD;
	T :	TIME;

	Y :	DWORD;

	func_block : FILTER_DW;
  END_VAR
	func_block.X  := X;
	func_block.T  := T;
	func_block();
	Y := func_block.Y;
END_PROGRAM

CONFIGURATION Config0
	VAR_GLOBAL
		PLC_TICKS_PER_SEC :	INT;
		PLC_SYS_TICK_CNT :	DINT;
	END_VAR
	RESOURCE Res0 ON PLC
		TASK task0(INTERVAL := T#20ms,PRIORITY := 0);
		PROGRAM instance0 WITH task0 : program0;
	END_RESOURCE
END_CONFIGURATION

(* ---- 563-HTML_ENCODE.ST ---- *)
FUNCTION_BLOCK HTML_ENCODE

	VAR_INPUT
		IN :	oscat_STRING250;
		M :	BOOL;
	END_VAR

	VAR_OUTPUT
		HTML_ENCODE :	oscat_STRING250;
	END_VAR

	VAR
		pt_out :	oscat_aB1_255;
		pos_in :	INT;
		pos_out :	INT;
		stop :	INT;
		B :	INT;
		tmp :	oscat_STRING10;
		i :	INT;
		BUF_TO_STRING :	BUF_TO_STRING;
		CHARNAME :	CHARNAME;
		CODE :	CODE;
	END_VAR

	pos_in := 1;
	stop := LEN(in);
	FOR pos_out := 1 TO 250 DO
		IF pos_in > stop THEN EXIT; END_IF;
		B := GET_CHAR(IN,pos_in);
		CASE B OF
			34:
				IF pos_out > 244 THEN EXIT; END_IF;
				pt_out[pos_out] := BYTE#38;
				pos_out := pos_out + 1;
				pt_out[pos_out] := BYTE#113;
				pos_out := pos_out + 1;
				pt_out[pos_out] := BYTE#117;
				pos_out := pos_out + 1;
				pt_out[pos_out] := BYTE#111;
				pos_out := pos_out + 1;
				pt_out[pos_out] := BYTE#116;
				pos_out := pos_out + 1;
				pt_out[pos_out] := BYTE#59;
			38:
				IF pos_out > 245 THEN EXIT; END_IF;
				pt_out[pos_out] := BYTE#38;
				pos_out := pos_out + 1;
				pt_out[pos_out] := BYTE#97;
				pos_out := pos_out + 1;
				pt_out[pos_out] := BYTE#109;
				pos_out := pos_out + 1;
				pt_out[pos_out] := BYTE#112;
				pos_out := pos_out + 1;
				pt_out[pos_out] := BYTE#59;
			60:
				IF pos_out > 246 THEN EXIT; END_IF;
				pt_out[pos_out] := BYTE#38;
				pos_out := pos_out + 1;
				pt_out[pos_out] := BYTE#108;
				pos_out := pos_out + 1;
				pt_out[pos_out] := BYTE#116;
				pos_out := pos_out + 1;
				pt_out[pos_out] := BYTE#59;
			62:
				IF pos_out > 246 THEN EXIT; END_IF;
				pt_out[pos_out] := BYTE#38;
				pos_out := pos_out + 1;
				pt_out[pos_out] := BYTE#103;
				pos_out := pos_out + 1;
				pt_out[pos_out] := BYTE#116;
				pos_out := pos_out + 1;
				pt_out[pos_out] := BYTE#59;
		ELSE
			IF M AND B > 127 THEN
				CHARNAME(C:=INT_TO_BYTE(B));
				tmp := CHARNAME.CHARNAME;
				IF pos_out + LEN(tmp) + 2 <= 250 THEN
					pt_out[pos_out] := BYTE#38;
					pos_out := pos_out + 1;
					FOR i := 1 TO LEN(tmp) DO
						CODE(STR:=tmp,POS:=i);
						pt_out[pos_out] := CODE.CODE;
						pos_out := pos_out + 1;
					END_FOR;
					pt_out[pos_out] := BYTE#59;
				END_IF;
			ELSE
			pt_out[pos_out] := INT_TO_BYTE(B);
			END_IF;
		END_CASE;
		pos_in := pos_in + 1;
	END_FOR;

	pos_out := pos_out - 1;

	FOR pos_in := 0 TO 1 DO
	BUF_TO_STRING.REQ        := pos_in>0;
	BUF_TO_STRING.BUF_FORMAT := TRUE;
	BUF_TO_STRING.BUF_OFFS   := DINT#0;
	BUF_TO_STRING.BUF_CNT    := INT_TO_DINT(pos_out);
	BUF_TO_STRING.BUFFER     := pt_out;
	BUF_TO_STRING.DST        := HTML_ENCODE;
	BUF_TO_STRING();
	pt_out  := BUF_TO_STRING.BUFFER;
	HTML_ENCODE := BUF_TO_STRING.DST;
	END_FOR;

END_FUNCTION_BLOCK

(* ---- 565-ESR_COLLECT.ST ---- *)
TYPE
	oscat_esr_collect_data      : ARRAY [0..7]    OF BYTE;
END_TYPE
TYPE oscat_esr_data :
  STRUCT
	typ    : BYTE;
	adress : STRING;
	DS     : UDINT;
	TS     : TIME;
	data   : oscat_esr_collect_data;
  END_STRUCT;
END_TYPE

TYPE
  oscat_ESR_3                : ARRAY [0..3] OF oscat_esr_data;
  oscat_ESR_31               : ARRAY [0..31] OF oscat_esr_data;
END_TYPE

FUNCTION INC1:INT

	VAR_INPUT
		X :	INT;
		N :	INT;
	END_VAR

	IF X >= N - 1 THEN
		INC1 := 0;
	ELSE
		INC1 := X + 1;
	END_IF;
END_FUNCTION

FUNCTION_BLOCK ESR_COLLECT
	VAR_INPUT
		ESR_0 :	oscat_ESR_3;
		ESR_1 :	oscat_ESR_3;
		ESR_2 :	oscat_ESR_3;
		ESR_3 :	oscat_ESR_3;
		ESR_4 :	oscat_ESR_3;
		ESR_5 :	oscat_ESR_3;
		ESR_6 :	oscat_ESR_3;
		ESR_7 :	oscat_ESR_3;
		RST :	BOOL;
	END_VAR

	VAR_IN_OUT
		POS :	INT;
	END_VAR

	VAR_OUTPUT
		ESR_OUT :	oscat_ESR_31;
	END_VAR

	VAR
		cnt :	INT := -1;
		max_in :	INT := 3;
		max_out :	INT := 32;
	END_VAR

	IF rst OR cnt < 0 THEN
		pos := -1;
	ELSE
		FOR cnt := 0 TO max_in DO
		IF esr_0[cnt].typ > BYTE#0 THEN pos := INC1(pos, max_out); esr_out[pos] := esr_0[cnt]; END_IF;
		IF esr_1[cnt].typ > BYTE#0 THEN pos := INC1(pos, max_out); esr_out[pos] := esr_1[cnt]; END_IF;
		IF esr_2[cnt].typ > BYTE#0 THEN pos := INC1(pos, max_out); esr_out[pos] := esr_2[cnt]; END_IF;
		IF esr_3[cnt].typ > BYTE#0 THEN pos := INC1(pos, max_out); esr_out[pos] := esr_3[cnt]; END_IF;
		IF esr_4[cnt].typ > BYTE#0 THEN pos := INC1(pos, max_out); esr_out[pos] := esr_4[cnt]; END_IF;
		IF esr_5[cnt].typ > BYTE#0 THEN pos := INC1(pos, max_out); esr_out[pos] := esr_5[cnt]; END_IF;
		IF esr_6[cnt].typ > BYTE#0 THEN pos := INC1(pos, max_out); esr_out[pos] := esr_6[cnt]; END_IF;
		IF esr_7[cnt].typ > BYTE#0 THEN pos := INC1(pos, max_out); esr_out[pos] := esr_7[cnt]; END_IF;
	END_FOR;
	END_IF;

END_FUNCTION_BLOCK

PROGRAM program0
  VAR
	ESR_0 :	oscat_ESR_3;
	ESR_1 :	oscat_ESR_3;
	ESR_2 :	oscat_ESR_3;
	ESR_3 :	oscat_ESR_3;
	ESR_4 :	oscat_ESR_3;
	ESR_5 :	oscat_ESR_3;
	ESR_6 :	oscat_ESR_3;
	ESR_7 :	oscat_ESR_3;
	RST   :	BOOL;

	POS   :	INT;

	ESR_OUT :	oscat_ESR_31;

	func_block : ESR_COLLECT;
  END_VAR
	func_block.ESR_0 :=ESR_0;
	func_block.ESR_1 :=ESR_1;
	func_block.ESR_2 :=ESR_2;
	func_block.ESR_3 :=ESR_3;
	func_block.ESR_4 :=ESR_4;
	func_block.ESR_5 :=ESR_5;
	func_block.ESR_6 :=ESR_6;
	func_block.ESR_7 :=ESR_7;
	func_block.RST   :=RST  ;
	func_block.POS   :=POS  ;

	func_block();
	POS := func_block.POS;
	ESR_OUT := func_block.ESR_OUT;

END_PROGRAM

CONFIGURATION Config0
	RESOURCE Res0 ON PLC
		TASK task0(INTERVAL := T#20ms,PRIORITY := 0);
		PROGRAM instance0 WITH task0 : program0;
	END_RESOURCE
END_CONFIGURATION

(* ---- 566-FLOAT_TO_REAL.ST ---- *)
FUNCTION BIT_OF_DWORD : BOOL
  VAR_INPUT
    IN : DWORD;
    N : INT;
  END_VAR

  BIT_OF_DWORD := (SHR(in,N) AND 16#00000001) > 0;
END_FUNCTION

FUNCTION EXPN:REAL

	VAR_INPUT
		X :	REAL;
		N :	INT;
	END_VAR

	VAR
		N_word :	WORD;
		X_tmp :	REAL;
		sign :	BOOL;
	END_VAR

	N_word := INT_TO_WORD(N);
	X_tmp := X;
	sign := BIT_OF_DWORD(WORD_TO_DWORD(N_word),15);
	N_word := INT_TO_WORD(ABS(N));
	IF BIT_OF_DWORD(WORD_TO_DWORD(N_word),0) THEN expn := X_tmp; ELSE expn := 1.0; END_IF;    (* N_word.X0 *)
	N_word := SHR(N_word,1);
	WHILE N_word > WORD#0 DO
		X_tmp := X_tmp * X_tmp;
		IF BIT_OF_DWORD(WORD_TO_DWORD(N_word),0) THEN expn := expn * X_tmp; END_IF;       (* N_word.X0 *)
		N_word := SHR(N_word,1);
	END_WHILE;
	IF sign THEN EXPN := 1.0 / EXPN; END_IF;

END_FUNCTION

FUNCTION_BLOCK FLOAT_TO_REAL_Block

	VAR_INPUT
		FLT :	STRING;
	END_VAR

	VAR_OUTPUT
		FLOAT_TO_REAL :	REAL;
	END_VAR

	VAR
		i :	INT;
		X :	BYTE;
		sign :	INT := 1;
		stop :	INT;
		tmp :	DINT;
		d :	INT;
		DEC_TO_INT :	DEC_TO_INT;
		CODE :	CODE;
	END_VAR

	sign := 1;
	d := 0;
	stop := LEN(FLT);
	tmp := DINT#0;

	FOR i := 1 TO stop DO
		CODE(STR:=FLT,POS:=i);
		X := CODE.CODE;
		IF X > BYTE#47 AND X < BYTE#58 OR X = BYTE#46 THEN
			EXIT;
		ELSIF X = BYTE#45 THEN
			(* code 45 is sign *)
			sign := -1;
		END_IF;
	END_FOR;

	FOR i := i TO stop DO
		CODE(STR:=FLT,POS:=i);
		X := CODE.CODE;
		IF X = BYTE#44 OR X = BYTE#46 OR X = BYTE#69 OR X = BYTE#101 THEN
			EXIT;
		(* calculate the value of the digit *)
		ELSIF X > BYTE#47 AND x < BYTE#58 THEN
			tmp := tmp * DINT#10 + _BYTE_TO_DINT(X) - DINT#48;
		END_IF;
	END_FOR;

	IF x = BYTE#44 OR X = BYTE#46 THEN
		FOR i := i + 1 TO stop DO
			CODE(STR:=FLT,POS:=i);
			X := CODE.CODE;
			IF X = BYTE#69 OR X = BYTE#101 THEN
				EXIT;
			ELSIF x > BYTE#47 AND x < BYTE#58 THEN
				tmp := tmp * DINT#10 + _BYTE_TO_DINT(X) - DINT#48;
				d := d - 1;
			END_IF;
		END_FOR;
	END_IF;

	IF (X = BYTE#69 OR X = BYTE#101) AND i<=stop THEN
		DEC_TO_INT(DEC:=MID(FLT, MIN(stop - i,10),MIN(stop,i+1)));
		d := d + DEC_TO_INT.DEC_TO_INT;

	(*    DEC_TO_INT(DEC:=RIGHT(FLT, MIN(stop - i,10)));
		d := d + DEC_TO_INT.DEC_TO_INT;*)
	END_IF;

	FLOAT_TO_REAL :=  EXPN(10.0, d) * DINT_TO_REAL(TMP * INT_TO_DINT(SIGN));

END_FUNCTION_BLOCK

PROGRAM program0
  VAR
    LocalVar0 : STRING;
	LocalOUT  : REAL;
	func_block : FLOAT_TO_REAL_Block;
  END_VAR
	func_block.FLT  := LocalVar0;
	func_block();
	LocalOUT := func_block.FLOAT_TO_REAL;
END_PROGRAM

CONFIGURATION Config0
  RESOURCE Res0 ON PLC
    TASK task0(INTERVAL := T#20ms,PRIORITY := 0);
    PROGRAM instance0 WITH task0 : program0;
  END_RESOURCE
END_CONFIGURATION

(* ---- 568-SETUP_HOLIDAY_FR.ST ---- *)
TYPE oscat_HOLIDAY_DATA :
	STRUCT
		NAME : STRING;
		DAY : SINT;
		MONTH : SINT;
		USE : SINT;
		PAD_BYTE : BYTE;
	END_STRUCT;
END_TYPE

TYPE
	oscat_HOLIDAY_DATA_0_29 	: ARRAY [0..29] OF oscat_HOLIDAY_DATA;
END_TYPE

FUNCTION_BLOCK SETUP_HOLIDAY_FR_Block

	VAR_IN_OUT
		HD :	oscat_HOLIDAY_DATA_0_29;
	END_VAR

	VAR
		init :	BOOL;
	END_VAR

	IF init THEN RETURN; END_IF;

	init := TRUE;

	HD[00].NAME := 'Nouve an';
	HD[00].DAY  := SINT#01;
	HD[00].MONTH := SINT#01;
	HD[00].USE := SINT#01;

	HD[01].NAME := 'St Valentin';
	HD[01].DAY  := SINT#14;
	HD[01].MONTH := SINT#02;
	HD[01].USE := SINT#00;

	HD[02].NAME := 'Vendredi Saint (alsace)';
	HD[02].DAY  := SINT#-2;
	HD[02].MONTH := SINT#00;
	HD[02].USE := SINT#00;

	HD[03].NAME := 'Dimanche de pques';
	HD[03].DAY  := SINT#00;
	HD[03].MONTH := SINT#00;
	HD[03].USE := SINT#01;

	HD[04].NAME := 'Lundi de pques';
	HD[04].DAY  := SINT#01;
	HD[04].MONTH := SINT#00;
	HD[04].USE := SINT#01;

	HD[05].NAME := 'Jeudi de Ascension';
	HD[05].DAY  := SINT#39;
	HD[05].MONTH := SINT#00;
	HD[05].USE := SINT#01;

	HD[06].NAME := 'dimanche de Pentecte';
	HD[06].DAY  := SINT#49;
	HD[06].MONTH := SINT#00;
	HD[06].USE := SINT#01;

	HD[07].NAME := 'jeudi de la Trinit';
	HD[07].DAY  := SINT#60;
	HD[07].MONTH := SINT#00;
	HD[07].USE := SINT#00;

	HD[08].NAME := 'Fte du travail';
	HD[08].DAY  := SINT#01;
	HD[08].MONTH := SINT#05;
	HD[08].USE := SINT#01;

	HD[09].NAME := 'Victoire 1945 ';
	HD[09].DAY  := SINT#08;
	HD[09].MONTH := SINT#05;
	HD[09].USE := SINT#01;

	HD[10].NAME := 'Prise de La bastille';
	HD[10].DAY  := SINT#14;
	HD[10].MONTH := SINT#07;
	HD[10].USE := SINT#01;

	HD[11].NAME := '15 Aot 1944';
	HD[11].DAY  := SINT#15;
	HD[11].MONTH := SINT#08;
	HD[11].USE := SINT#01;

	HD[12].NAME := 'Halloween';
	HD[12].DAY  := SINT#31;
	HD[12].MONTH := SINT#10;
	HD[12].USE := SINT#00;

	HD[13].NAME := 'Armistice 1918';
	HD[13].DAY  := SINT#11;
	HD[13].MONTH := SINT#11;
	HD[13].USE := SINT#01;

	HD[14].NAME := 'Nol';
	HD[14].DAY  := SINT#25;
	HD[14].MONTH := SINT#12;
	HD[14].USE := SINT#01;

	HD[15].NAME := 'Saint tienne (alsace)';
	HD[15].DAY  := SINT#26;
	HD[15].MONTH := SINT#12;
	HD[15].USE := SINT#00;

	HD[16].NAME := 'Fte de la musique';
	HD[16].DAY  := SINT#21;
	HD[16].MONTH := SINT#06;
	HD[16].USE := SINT#00;
END_FUNCTION_BLOCK

PROGRAM program0
  VAR
    LocalVar0 : oscat_HOLIDAY_DATA_0_29;
	func_block : SETUP_HOLIDAY_FR_Block;
  END_VAR
	func_block.HD  := LocalVar0;
	func_block();
	LocalVar0 := func_block.HD;
END_PROGRAM

CONFIGURATION Config0
  RESOURCE Res0 ON PLC
    TASK task0(INTERVAL := T#20ms,PRIORITY := 0);
    PROGRAM instance0 WITH task0 : program0;
  END_RESOURCE
END_CONFIGURATION

(* ---- 569-SIGNAL.ST ---- *)
FUNCTION _BYTE_TO_INT:INT
	VAR_INPUT
		IN :	BYTE;
	END_VAR

	_BYTE_TO_INT := USINT_TO_INT(BYTE_TO_USINT(IN));
END_FUNCTION

FUNCTION TIME_TO_UDINT2:UDINT
	VAR_INPUT
		X :	TIME;
	END_VAR

	TIME_TO_UDINT2 := DINT_TO_UDINT(TIME_TO_DINT(X));
END_FUNCTION

FUNCTION UDINT_TO_TIME2:TIME

	VAR_INPUT
		IN :	UDINT;
	END_VAR

	UDINT_TO_TIME2 := DINT_TO_TIME(UDINT_TO_DINT(IN));

END_FUNCTION

FUNCTION_BLOCK T_PLC_MS_block
	VAR_OUTPUT
		T_PLC_MS :	UDINT;
	END_VAR

	VAR_EXTERNAL
		PLC_TICKS_PER_SEC :	INT;
		PLC_SYS_TICK_CNT :	DINT;
	END_VAR

	VAR
		debug :	BOOL;(*Debug-Mode ON / OFF*)
		N :	INT;(*Debug-Faktor*)
		Offset :	UDINT;(*Debug-Offset*)
		temp :	DWORD := DWORD#1;(*Debug-Offset*)
		mode :	BOOL;(*modus*)
		faktor :	UDINT;(*Systemtakt-Faktor*)
		init :	BOOL;
		v_plc_ticks_per_sec :	UDINT;
		base :	UDINT := UDINT#1000;
	END_VAR

	IF init = FALSE THEN
		v_plc_ticks_per_sec := INT_TO_UDINT(PLC_TICKS_PER_SEC);
		IF v_plc_ticks_per_sec = UDINT#1024 THEN
			faktor := UDINT#1;
			mode := FALSE;
		ELSIF v_plc_ticks_per_sec > UDINT#0 THEN
			IF v_plc_ticks_per_sec <= base THEN
				faktor := base / v_plc_ticks_per_sec;
				mode := FALSE;
			ELSE
				faktor := v_plc_ticks_per_sec / base;
				mode := TRUE;
			END_IF;
		ELSE
			faktor := UDINT#1;
		END_IF;
		init := TRUE;
	END_IF;

	IF mode THEN
		T_PLC_MS := DINT_TO_UDINT(PLC_SYS_TICK_CNT) / faktor;
	ELSE
		T_PLC_MS := DINT_TO_UDINT(PLC_SYS_TICK_CNT) * faktor;
	END_IF;

	IF debug THEN
		T_PLC_MS := (DWORD_TO_UDINT(SHL(UDINT_TO_DWORD(T_PLC_MS),N) OR SHL(temp,N)) - UDINT#1) + Offset;
	END_IF;

END_FUNCTION_BLOCK

FUNCTION_BLOCK SIGNAL_Block

	VAR_INPUT
		IN :	BOOL;
		SIG :	BYTE;
		TS :	TIME;
	END_VAR

	VAR_OUTPUT
		Q :	BOOL;
	END_VAR

	VAR
		tx :	DWORD;
		_step :	BYTE;
		T_PLC_MS :	T_PLC_MS_Block;
	END_VAR

	IF in THEN
		T_PLC_MS();
		tx:= UDINT_TO_DWORD(T_PLC_MS.T_PLC_MS);

		IF ts > t#0s THEN
			_step := DWORD_TO_BYTE(UDINT_TO_DWORD(DWORD_TO_UDINT(tx) / TIME_TO_UDINT2(ts)) AND DWORD#16#0000_0007);
		ELSE
			_step := DWORD_TO_BYTE(SHR(tx,7) AND DWORD#16#0000_0007);
		END_IF;
		_step := SHL(BYTE#1,_BYTE_TO_INT(_step));
		Q := (_step AND sig) > BYTE#0;
	ELSE
		Q := FALSE;
	END_IF;

END_FUNCTION_BLOCK

PROGRAM program0
  VAR
	IN :	BOOL;
	SIG :	BYTE;
	TS :	TIME;
	Q :	BOOL;
	func_block : SIGNAL_Block;
  END_VAR
	func_block.IN  :=IN;
	func_block.SIG  :=SIG;
	func_block.TS  :=TS;
	func_block();
	Q := func_block.Q;

END_PROGRAM

CONFIGURATION Config0

	VAR_GLOBAL
		PLC_TICKS_PER_SEC :	INT;
		PLC_SYS_TICK_CNT :	DINT;
	END_VAR

  	RESOURCE Res0 ON PLC
    	TASK task0(INTERVAL := T#20ms,PRIORITY := 0);
    	PROGRAM instance0 WITH task0 : program0;
  	END_RESOURCE

END_CONFIGURATION

(* ---- 570-DT_SIMU.ST ---- *)
FUNCTION _REAL_TO_UDINT:UDINT
  VAR_INPUT
    X :	REAL;
  END_VAR

  IF REAL_TO_UDINT(0.5) = UDINT#1 THEN
    _REAL_TO_UDINT := REAL_TO_UDINT(x);
  ELSIF X > 0.0 THEN
    _REAL_TO_UDINT := REAL_TO_UDINT(x+0.5);
  ELSIF X < 0.0 THEN
    _REAL_TO_UDINT := REAL_TO_UDINT(x-0.5);
  ELSE
    _REAL_TO_UDINT := UDINT#0;
  END_IF;
END_FUNCTION

FUNCTION_BLOCK T_PLC_MS_block

	VAR_OUTPUT
		T_PLC_MS :	UDINT;
	END_VAR

	VAR_EXTERNAL
		PLC_TICKS_PER_SEC :	INT;
		PLC_SYS_TICK_CNT :	DINT;
	END_VAR

	VAR
		debug :	BOOL;(*Debug-Mode ON / OFF*)
		N :	INT;(*Debug-Faktor*)
		Offset :	UDINT;(*Debug-Offset*)
		temp :	DWORD := DWORD#1;(*Debug-Offset*)
		mode :	BOOL;(*modus*)
		faktor :	UDINT;(*Systemtakt-Faktor*)
		init :	BOOL;
		v_plc_ticks_per_sec :	UDINT;
		base :	UDINT := UDINT#1000;
	END_VAR

	IF init = FALSE THEN
		v_plc_ticks_per_sec := INT_TO_UDINT(PLC_TICKS_PER_SEC);
		IF v_plc_ticks_per_sec = UDINT#1024 THEN
			faktor := UDINT#1;
			mode := FALSE;
		ELSIF v_plc_ticks_per_sec > UDINT#0 THEN
			IF v_plc_ticks_per_sec <= base THEN
				faktor := base / v_plc_ticks_per_sec;
				mode := FALSE;
			ELSE
				faktor := v_plc_ticks_per_sec / base;
				mode := TRUE;
			END_IF;
		ELSE
			faktor := UDINT#1;
		END_IF;
		init := TRUE;
	END_IF;

	IF mode THEN
		T_PLC_MS := DINT_TO_UDINT(PLC_SYS_TICK_CNT) / faktor;
	ELSE
		T_PLC_MS := DINT_TO_UDINT(PLC_SYS_TICK_CNT) * faktor;
	END_IF;

	IF debug THEN
		T_PLC_MS := (DWORD_TO_UDINT(SHL(UDINT_TO_DWORD(T_PLC_MS),N) OR SHL(temp,N)) - UDINT#1) + Offset;
	END_IF;

END_FUNCTION_BLOCK

FUNCTION_BLOCK DT_SIMU
	VAR_INPUT
		START :	UDINT;
		SPEED :	REAL := 1.0;
	END_VAR

	VAR_OUTPUT
		DTS :	UDINT;
	END_VAR

	VAR
		tc :	UDINT;
		init :	BOOL;
		last :	UDINT;
		tx :	UDINT;
		td :	UDINT;
		T_PLC_MS :	T_PLC_MS_block;
	END_VAR

	T_PLC_MS();
	tx:= T_PLC_MS.T_PLC_MS;
	tc := _REAL_TO_UDINT(UDINT_TO_REAL(tx - last) * speed);

	IF NOT init THEN
		init := TRUE;
		DTS := Start;
		tc := UDINT#0;
		last := tx;
	ELSIF SPEED = 0.0 THEN
		DTS := DTS + UDINT#1;
	ELSIF tc >= UDINT#1000 THEN
		td := (tc / UDINT#1000) * UDINT#1000;
		DTS := DTS + td;
		last := last + _REAL_TO_UDINT(UDINT_TO_REAL(td) / speed);
	END_IF;
END_FUNCTION_BLOCK

PROGRAM program0
  VAR
    LocalVar0 : UDINT;
	LocalVar1 : REAL;
	LocalOUT  : UDINT;
	func_block : DT_SIMU;
  END_VAR
	func_block.START  := LocalVar0;
	func_block.SPEED  := LocalVar1;
	func_block();
	LocalOUT := func_block.DTS;
END_PROGRAM

CONFIGURATION Config0

	VAR_GLOBAL
		PLC_TICKS_PER_SEC :	INT;
		PLC_SYS_TICK_CNT :	DINT;
	END_VAR

  	RESOURCE Res0 ON PLC
    	TASK task0(INTERVAL := T#20ms,PRIORITY := 0);
    	PROGRAM instance0 WITH task0 : program0;
  	END_RESOURCE

END_CONFIGURATION

(* ---- 571-FT_RMP.ST ---- *)
FUNCTION_BLOCK T_PLC_MS_block
	VAR_OUTPUT
		T_PLC_MS :	UDINT;
	END_VAR

	VAR_EXTERNAL
		PLC_TICKS_PER_SEC :	INT;
		PLC_SYS_TICK_CNT :	DINT;
	END_VAR

	VAR
		debug :	BOOL;(*Debug-Mode ON / OFF*)
		N :	INT;(*Debug-Faktor*)
		Offset :	UDINT;(*Debug-Offset*)
		temp :	DWORD := DWORD#1;(*Debug-Offset*)
		mode :	BOOL;(*modus*)
		faktor :	UDINT;(*Systemtakt-Faktor*)
		init :	BOOL;
		v_plc_ticks_per_sec :	UDINT;
		base :	UDINT := UDINT#1000;
	END_VAR

	IF init = FALSE THEN
		v_plc_ticks_per_sec := INT_TO_UDINT(PLC_TICKS_PER_SEC);
		IF v_plc_ticks_per_sec = UDINT#1024 THEN
			faktor := UDINT#1;
			mode := FALSE;
		ELSIF v_plc_ticks_per_sec > UDINT#0 THEN
			IF v_plc_ticks_per_sec <= base THEN
				faktor := base / v_plc_ticks_per_sec;
				mode := FALSE;
			ELSE
				faktor := v_plc_ticks_per_sec / base;
				mode := TRUE;
			END_IF;
		ELSE
			faktor := UDINT#1;
		END_IF;
		init := TRUE;
	END_IF;

	IF mode THEN
		T_PLC_MS := DINT_TO_UDINT(PLC_SYS_TICK_CNT) / faktor;
	ELSE
		T_PLC_MS := DINT_TO_UDINT(PLC_SYS_TICK_CNT) * faktor;
	END_IF;

	IF debug THEN
		T_PLC_MS := (DWORD_TO_UDINT(SHL(UDINT_TO_DWORD(T_PLC_MS),N) OR SHL(temp,N)) - UDINT#1) + Offset;
	END_IF;
END_FUNCTION_BLOCK

FUNCTION_BLOCK FT_RMP

	VAR_INPUT
		RMP :	BOOL := TRUE;
		IN :	REAL;
		KR :	REAL;
		KF :	REAL;
	END_VAR

	VAR_OUTPUT
		OUT :	REAL;
		BUSY :	BOOL;
		UD :	BOOL;
	END_VAR

	VAR
		tx :	TIME;
		last :	TIME;
		init :	BOOL;
		T_PLC_MS :	T_PLC_MS_block;
	END_VAR

	T_PLC_MS();
	tx:= UDINT_TO_TIME(T_PLC_MS.T_PLC_MS) - last;

	IF NOT init THEN
		init := TRUE;
		last := tx;
		tx := t#0s;
		out := in;
	END_IF;
	IF NOT rmp THEN
		out := in;
		busy := FALSE;
	ELSIF out > in THEN
		(* ramp down *)
		out := out - TIME_TO_REAL(tx) * 0.001 * KF;
		out := MAX(in, out);
	ELSIF out < in THEN
		(* ramp up *)
		out := out + TIME_TO_REAL(tx) * 0.001 * KR;
		out := MIN(in, out);
	END_IF;

	(* set busy and dir flags *)
	IF out < in THEN
		busy := TRUE;
		ud := TRUE;
	ELSIF out > in THEN
		busy := TRUE;
		ud := FALSE;
	ELSE
		busy := FALSE;
	END_IF;
	last := last + tx;

END_FUNCTION_BLOCK

PROGRAM program0
	VAR
		RMP :	BOOL := TRUE;
		IN :	REAL;
		KR :	REAL;
		KF :	REAL;

		OUT :	REAL;
		BUSY :	BOOL;
		UD :	BOOL;

		func_block : FT_RMP;
	END_VAR
	func_block.RMP := RMP;
	func_block.IN := IN;
	func_block.KR := KR;
	func_block.KF := KF;
	func_block();
	OUT := func_block.OUT;
	BUSY := func_block.BUSY;
	UD := func_block.UD;

END_PROGRAM

CONFIGURATION Config0

	VAR_GLOBAL
		PLC_TICKS_PER_SEC :	INT;
		PLC_SYS_TICK_CNT :	DINT;
	END_VAR

	RESOURCE Res0 ON PLC
		TASK task0(INTERVAL := T#20ms,PRIORITY := 0);
		PROGRAM instance0 WITH task0 : program0;
	END_RESOURCE

END_CONFIGURATION

(* ---- 572-PULSE_LENGTH.ST ---- *)
FUNCTION UDINT_TO_TIME2:TIME

	VAR_INPUT
		IN :	UDINT;
	END_VAR

	UDINT_TO_TIME2 := DINT_TO_TIME(UDINT_TO_DINT(IN));

END_FUNCTION

FUNCTION_BLOCK T_PLC_MS_block
	VAR_OUTPUT
		T_PLC_MS :	UDINT;
	END_VAR

	VAR_EXTERNAL
		PLC_TICKS_PER_SEC :	INT;
		PLC_SYS_TICK_CNT :	DINT;
	END_VAR

	VAR
		debug :	BOOL;(*Debug-Mode ON / OFF*)
		N :	INT;(*Debug-Faktor*)
		Offset :	UDINT;(*Debug-Offset*)
		temp :	DWORD := DWORD#1;(*Debug-Offset*)
		mode :	BOOL;(*modus*)
		faktor :	UDINT;(*Systemtakt-Faktor*)
		init :	BOOL;
		v_plc_ticks_per_sec :	UDINT;
		base :	UDINT := UDINT#1000;
	END_VAR

	IF init = FALSE THEN
		v_plc_ticks_per_sec := INT_TO_UDINT(PLC_TICKS_PER_SEC);
		IF v_plc_ticks_per_sec = UDINT#1024 THEN
			faktor := UDINT#1;
			mode := FALSE;
		ELSIF v_plc_ticks_per_sec > UDINT#0 THEN
			IF v_plc_ticks_per_sec <= base THEN
				faktor := base / v_plc_ticks_per_sec;
				mode := FALSE;
			ELSE
				faktor := v_plc_ticks_per_sec / base;
				mode := TRUE;
			END_IF;
		ELSE
			faktor := UDINT#1;
		END_IF;
		init := TRUE;
	END_IF;

	IF mode THEN
		T_PLC_MS := DINT_TO_UDINT(PLC_SYS_TICK_CNT) / faktor;
	ELSE
		T_PLC_MS := DINT_TO_UDINT(PLC_SYS_TICK_CNT) * faktor;
	END_IF;

	IF debug THEN
		T_PLC_MS := (DWORD_TO_UDINT(SHL(UDINT_TO_DWORD(T_PLC_MS),N) OR SHL(temp,N)) - UDINT#1) + Offset;
	END_IF;

END_FUNCTION_BLOCK

FUNCTION_BLOCK PULSE_LENGTH_Block

	VAR_INPUT
		IN :	BOOL;
		T_SHORT :	TIME := T#100ms;
		T_LONG :	TIME := T#1s;
	END_VAR

	VAR_OUTPUT
		SHORT :	BOOL;
		MIDDLE :	BOOL;
		LONG :	BOOL;
	END_VAR

	VAR
		tx :	TIME;
		tn :	TIME;
		edge :	BOOL;
		T_PLC_MS :	T_PLC_MS_Block;
	END_VAR

	T_PLC_MS();
	tx:= UDINT_TO_TIME(T_PLC_MS.T_PLC_MS);

	short := FALSE;
	Middle := FALSE;
	long := FALSE;

	IF in AND NOT edge THEN
		edge := TRUE;
		tn := tx;

	ELSIF NOT in AND edge THEN
		edge := FALSE;
		tn := tx - tn;
		IF tn < t_short THEN
			short := TRUE;
		ELSIF tn > t_long THEN
			long := TRUE;
		ELSE
			Middle := TRUE;
		END_IF;

	ELSIF in AND tx - tn > t_long THEN
		long := TRUE;
	END_IF;

END_FUNCTION_BLOCK

PROGRAM program0
	VAR
		IN :	BOOL;
		T_SHORT :	TIME := T#100ms;
		T_LONG :	TIME := T#1s;
		SHORT :	BOOL;
		MIDDLE :	BOOL;
		LONG :	BOOL;

		func_block : PULSE_LENGTH_Block;
	END_VAR
	func_block.IN := IN;
	func_block.T_SHORT := T_SHORT;
	func_block.T_LONG := T_LONG ;

	func_block();
	SHORT  := func_block.SHORT;
	MIDDLE  := func_block.MIDDLE;
	LONG  := func_block.LONG;
END_PROGRAM

CONFIGURATION Config0
	VAR_GLOBAL
		PLC_TICKS_PER_SEC :	INT;
		PLC_SYS_TICK_CNT :	DINT;
	END_VAR
  	RESOURCE Res0 ON PLC
    	TASK task0(INTERVAL := T#20ms,PRIORITY := 0);
    	PROGRAM instance0 WITH task0 : program0;
  	END_RESOURCE
END_CONFIGURATION

(* ---- 573-TN_SC_FILL.ST ---- *)
TYPE
  bya_TN_CHAR:       	ARRAY [0..1919] OF BYTE;
  bya_TN_BACKUP:     	ARRAY [0..1919] OF BYTE;
  bya_TN_COLOR:      	ARRAY [0..1919] OF BYTE;
  bya_TN_Line_Update:	ARRAY [0..23]   OF BOOL;

  us_TN_SCREEN :
  STRUCT
		bya_CHAR:			bya_TN_CHAR;
		bya_COLOR:			bya_TN_COLOR;
		bya_BACKUP:			bya_TN_BACKUP;
		bya_Line_Update:	bya_TN_Line_Update;

		by_Input_Exten_Code:    BYTE;
		by_Input_ASCII_Code:    BYTE;
		bo_Input_ASCII_IsNum:   BOOL;
		in_Page_Number:        	INT;                (* aktive Seiten-Nr.              *)
		in_Cursor_X:           	INT;                (* Cursor X-Position              *)
		in_Cursor_Y:           	INT;                (* Cursor Y-Position              *)
		in_EOS_Offset:         	INT;                (* End of String Offset           *)
		by_Clear_Screen_Attr:  	BYTE;               (* Clear-Screen Attr              *)
		bo_Clear_Screen:       	BOOL;               (* Clear-Screen ausl�sen          *)
		bo_Modal_Dialog:       	BOOL;               (* Modaler Dialog ist aktiv       *)
		bo_Menue_Bar_Dialog:   	BOOL;               (* Menue Dialog ist aktiv         *)

  END_STRUCT;
END_TYPE

FUNCTION TN_SC_XY2_ERROR:BOOL

	VAR_INPUT
		X1 :	INT;
		Y1 :	INT;
		X2 :	INT;
		Y2 :	INT;
	END_VAR

	TN_SC_XY2_ERROR := Y1 < 0 OR X1 < 0 OR Y2 < 0 OR X2 < 0 OR Y1 > 23 OR X1 > 79 OR Y2 > 23 OR X2 > 79;

END_FUNCTION

FUNCTION_BLOCK TN_SC_FILL_Block

	VAR
		in_X :	INT;
		in_Y :	INT;
		in_Offset :	INT;
	END_VAR

	VAR_INPUT
		Iin_Y1 :	INT;
		Iin_X1 :	INT;
		Iin_Y2 :	INT;
		Iin_X2 :	INT;
		Iby_CHAR :	BYTE;
		Iby_Attr :	BYTE;
	END_VAR

	VAR_IN_OUT
		Xus_TN_SCREEN :	us_TN_SCREEN;
	END_VAR

	IF TN_SC_XY2_ERROR(Iin_X1,Iin_Y1,Iin_X2,Iin_Y2) THEN RETURN; END_IF;

	FOR in_Y := Iin_Y1 TO Iin_Y2 DO
	Xus_TN_SCREEN.bya_Line_Update[in_Y] := TRUE;
	in_Offset := (in_Y * 80) + Iin_X1;
	FOR in_X := Iin_X1 TO Iin_X2 DO
		Xus_TN_SCREEN.bya_CHAR[in_Offset]  := Iby_CHAR;
		Xus_TN_SCREEN.bya_COLOR[in_Offset] := Iby_Attr;
		in_Offset := in_Offset + 1;
	END_FOR;
	END_FOR;

END_FUNCTION_BLOCK

PROGRAM program0
	VAR
		Iin_Y1 :	INT;
		Iin_X1 :	INT;
		Iin_Y2 :	INT;
		Iin_X2 :	INT;
		Iby_CHAR :	BYTE;
		Iby_Attr :	BYTE;
		Xus_TN_SCREEN :	us_TN_SCREEN;

		func_block : TN_SC_FILL_Block;
	END_VAR
	func_block.Iin_X1 := Iin_X1;
	func_block.Iin_Y1 := Iin_Y1;
  	func_block.Iin_X2 := Iin_X2;
	func_block.Iin_Y2 := Iin_Y2;
  	func_block.Iby_CHAR := Iby_CHAR;
	func_block.Iby_Attr := Iby_Attr;
	func_block.Xus_TN_SCREEN := Xus_TN_SCREEN;

	func_block();
	Xus_TN_SCREEN  := func_block.Xus_TN_SCREEN;
END_PROGRAM

CONFIGURATION Config0
	RESOURCE Res0 ON PLC
		TASK task0(INTERVAL := T#20ms,PRIORITY := 0);
		PROGRAM instance0 WITH task0 : program0;
	END_RESOURCE
END_CONFIGURATION

(* ---- 575-M_D.ST ---- *)
FUNCTION_BLOCK T_PLC_MS_Block
	VAR_OUTPUT
		T_PLC_MS :	UDINT;
	END_VAR

	VAR_EXTERNAL
		PLC_TICKS_PER_SEC :	INT;
		PLC_SYS_TICK_CNT :	DINT;
	END_VAR

	VAR
		debug :	BOOL;(*Debug-Mode ON / OFF*)
		N :	INT;(*Debug-Faktor*)
		Offset :	UDINT;(*Debug-Offset*)
		temp :	DWORD := DWORD#1;(*Debug-Offset*)
		mode :	BOOL;(*modus*)
		faktor :	UDINT;(*Systemtakt-Faktor*)
		init :	BOOL;
		v_plc_ticks_per_sec :	UDINT;
		base :	UDINT := UDINT#1000;
	END_VAR

	IF init = FALSE THEN
		v_plc_ticks_per_sec := INT_TO_UDINT(PLC_TICKS_PER_SEC);
		IF v_plc_ticks_per_sec = UDINT#1024 THEN
			faktor := UDINT#1;
			mode := FALSE;
		ELSIF v_plc_ticks_per_sec > UDINT#0 THEN
			IF v_plc_ticks_per_sec <= base THEN
				faktor := base / v_plc_ticks_per_sec;
				mode := FALSE;
			ELSE
				faktor := v_plc_ticks_per_sec / base;
				mode := TRUE;
			END_IF;
		ELSE
			faktor := UDINT#1;
		END_IF;
		init := TRUE;
	END_IF;

	IF mode THEN
		T_PLC_MS := DINT_TO_UDINT(PLC_SYS_TICK_CNT) / faktor;
	ELSE
		T_PLC_MS := DINT_TO_UDINT(PLC_SYS_TICK_CNT) * faktor;
	END_IF;

	IF debug THEN
		T_PLC_MS := (DWORD_TO_UDINT(SHL(UDINT_TO_DWORD(T_PLC_MS),N) OR SHL(temp,N)) - UDINT#1) + Offset;
	END_IF;
END_FUNCTION_BLOCK

FUNCTION_BLOCK M_D_Block

	VAR_INPUT
		START :	BOOL;
		STOP :	BOOL;
		TMAX :	TIME := t#10d;
		RST :	BOOL;
	END_VAR

	VAR_OUTPUT
		PT :	TIME;
		ET :	TIME;
		RUN :	BOOL;
	END_VAR

	VAR
		edge :	BOOL;
		T0 :	TIME;
		tx :	TIME;
		startup :	BOOL;
		T_PLC_MS :	T_PLC_MS_Block;
	END_VAR

	(* check for rst input *)
	IF rst OR et >= tmax THEN
		pt := t#0ms;
		et := t#0ms;
		startup := FALSE;
		run := FALSE;
	END_IF;

	(* avoid timers to start when input is true at startup *)
	IF NOT startup THEN
		edge := start;
		startup := TRUE;
	END_IF;

	(* read system timer *)
	T_PLC_MS();
	tx:= UDINT_TO_TIME(T_PLC_MS.T_PLC_MS);

	(* detect rising edge on start *)
	IF start AND NOT edge AND NOT stop THEN
		t0 := tx;
		run := TRUE;
		pt := t#0s;
	ELSIF stop AND run THEN
		pt := et;
		run := FALSE;
	END_IF;
	edge := start;
	IF run THEN et := tx - t0; END_IF;

END_FUNCTION_BLOCK

PROGRAM program0

	VAR
		START :	BOOL;
		STOP :	BOOL;
		TMAX :	TIME := t#10d;
		RST :	BOOL;

		PT :	TIME;
		ET :	TIME;
		RUN :	BOOL;

		func_block : M_D_Block;
	END_VAR
	func_block.START := START;
	func_block.STOP := STOP;
	func_block.TMAX := TMAX;
	func_block.RST := RST;

	func_block();
	PT := func_block.PT;
	ET := func_block.ET;
	RUN := func_block.RUN;

END_PROGRAM

CONFIGURATION Config0

	VAR_GLOBAL
		PLC_TICKS_PER_SEC :	INT;
		PLC_SYS_TICK_CNT :	DINT;
	END_VAR

	RESOURCE Res0 ON PLC
		TASK task0(INTERVAL := T#20ms,PRIORITY := 0);
		PROGRAM instance0 WITH task0 : program0;
	END_RESOURCE

END_CONFIGURATION
